(* IEC 61131-3 sources: daoli-st-library/DL_Process (part 65) *)

(* ---- FB_DL_EnthalpyCompareCtrl.st ---- *)
(*==============================================================================
 * 组件名称 (Component)  : FB_DL_EnthalpyCompareCtrl
 * 所属子库 (Sublibrary) : DL_Process
 * 当前版本 (Version)    : 1.0.1
 * 组件分类 (Category)   : 功能块（FUNCTION_BLOCK）· 焓差经济器比较控制 ·
 *                         Level 2 行业池 9.5 节 P0 链路闭环示范
 * 兼容性   (Platform)   : CODESYS 3.5 / TwinCAT 3 / 汇川 InoProShop / Schneider
 *                         Machine Expert；仅依赖 Standard.library 与本库已入库
 *                         算法函数，零厂商方言
 * 功能描述 (Function)   : 焓差比较控制执行块。新风/回风温湿度 4 输入 → 每拍
 *                         两次调用 FC_DL_HumidAirEnthalpy 计算双侧比焓 →
 *                         差分焓值判据（施密特迟滞防临界抖动）→ 新风阀位指令
 *                         输出；含最小新风位硬下限（卫生通风底线）与 ASHRAE
 *                         90.1 新风焓值高限停机语义（回差=死区防振荡）。
 *
 * 【干球温度判据陷阱警示 / Dry-bulb trap warning】
 *   本块判据【只允许使用焓差】，严禁以干球温差（fOaTempC 与 fRaTempC 比较）
 *   代替焓差判据：湿工况下新风干球温度可以低于回风，但其潜热（含湿量）更高，
 *   总焓反而高于回风——若按干球降温直觉开大新风阀，会引入高焓湿空气增加表冷
 *   负荷（验收向量 V1 复现此陷阱）。任何把本块改为干球比较的改动均视为破坏
 *   焓差经济器物理语义。
 *
 * 设计要点 (Key notes)  : ① 连续量组件 → 设 bInit 首扫（R19 唯一合法范式
 *                           IF bTrack OR (NOT bInit)），首扫输出最小新风位
 *                           安全值并重建迟滞态，运行中途 bTrack 一拍即重同步；
 *                         ② 迟滞状态机：开侧 fOaEnth < fRaEnth − 死区、关侧
 *                           fOaEnth > fRaEnth + 死区，死区区间内保持原态
 *                           （传感器漂移防线）；CASE + ELSE 非法态兜底；
 *                         ③ 高限停机：fEnthalpyHighLimit > 0 使能，fOaEnth
 *                           ≥ 高限 → 停机锁 bHighLimitTrip，回落至
 *                           高限 − 死区 以下才解除（瞬时型每拍重算，R15）；
 *                         ④ 失效语义（R11 裁定 D2）：任一温湿度/大气压非有
 *                           限值或越出引脚域 → 阀位指令输出最小新风位（安全
 *                           侧兜底），fOaEnthalpy/fRaEnthalpy/bHighLimitTrip
 *                           冻结保持末次有效值（诊断量冻结），故障码锁存，
 *                           仅「输入恢复 + bReset 上升沿」解除（R15）；
 *                         ⑤ 时间/温湿度全部引脚注入，禁读 CPU 本地钟；
 *                         ⑥ 限幅域对调自修复：fMinOaPos > fFreeCoolOaPos
 *                           时对调继续计算（公约 0.6），量纲注释与限幅域一致。
 * 枚举归属 (Enum note)  : E_DL_EnthalpyHyst（迟滞双侧态）随本块同文件发布；
 *                         本块不重复声明任何既有枚举。
 * 依赖     (Depends)    : FC_DL_HumidAirEnthalpy（DL_Algo，公开接口直接调用，
 *                         不内联重实现其焓值公式）；Standard.library
 *                         （R_TRIG / ABS / MIN / MAX / LIMIT）。
 * 开源溯源 (Origin)     : 原创实现（参考 ASHRAE 90.1 economizer 高限判据与
 *                         OSCAT Building 焓差经济器行为定义，clean-room）。
 *                         仅借鉴公开判据语义（差分焓值切换、最小新风位底线、
 *                         高限停机），未读取、未复制任何源码行；迟滞状态机、
 *                         失效冻结语义与码表为本库独立设计。
 * 故障码表 (Error codes):
 *   16#0005_0202【故障级】焓值计算输入失效（非有限值/越引脚域，锁存，
 *                 解除条件：输入恢复 AND bReset 上升沿）
 *   16#0005_0201【故障级】非法状态兜底（CASE ELSE，复用本库既有同义码，
 *                 与 FB_DL_PackMlStateMachine 同语义，公共码先例
 *                 DL_Algo 16#0002_0004）
 *   16#0005_0103【信息级】下游算法函数钳位码透传归并（温度/湿度/大气压
 *                 越界已钳位照算）/ 限幅域对调自修复（公约 0.6，本块唯一
 *                 分配信息级码复用，见 R11 D3）
 * 【规格偏离留档 / R11 Deviation register】
 *   D1 规格分配故障码 0005_0201（输入失效）与子库既有台账冲突（0201 已被
 *      R5 PackML 非法状态兜底占用）：按公约 0.7 冲突顺延，输入失效改用
 *      0005_0202；非法状态兜底与规格 0005_0202 分配冲突 → 复用既有同义码
 *      0005_0201。语义不变，仅码位重排。
 *   D2 规格失效语义同时出现「冻结保持末次有效阀位」与「输出 fMinOaPos 兜
 *      底值」：裁定为阀位指令输出 fMinOaPos（安全侧），焓值诊断输出与高限
 *      锁存位冻结末次有效值。
 *   D3 限幅域对调自修复（公约 0.6）码位：本块仅分配信息级 0005_0103，对调
 *      事件与下游钳位透传共用该码（当拍 uErrorId 择一呈现，均为信息级）。
 *   D4 新风干球负温域（-30..0 摄氏度）超出下游焓值函数计算域（0..100）：
 *      负干球工况下游返回 0 摄氏度钳位焓值（对新风焓偏高估计 → 判据偏保守
 *      安全侧），钳位信息经 0005_0103 当拍呈现；是否放行负干球工况由调用方
 *      按 D4 取舍（本块按引脚域 -30..60 验收输入，不自行拒绝）。
 * 红线自检 (Redline)    : R1 ✓ 零全局变量表与外部变量引用 ｜ R2 ✓ 零物理 IO 地址直写
 *                         R3 ✓ 纯 IEC 61131-3 ｜ R4 ✓ 非有限值防御（fX<>fX 先检再比较）
 *                             +迟滞判据浮点禁判等+本块无除法运算
 *                         R5 ✓ 全变量中英双语同行注释 ｜ R6 ✓ 迟滞状态机 ENUM+CASE
 *                             且 CASE-ELSE 兜底（码 0005_0201）
 *                         R7 ✓ R_TRIG 实例主体无条件周期刷新（严禁入分支）
 * 修订历史 (Revision)   :
 *   2026-11-15  v1.0.0  首版入库 · Round 06 · 泳道 C · 契约出处 ROUND_PLAN_R6 §3.14
 *   2026-11-15  v1.0.1  终审修复【工程语义级】参数 REAL 输入非数防御缺口：
 *                       原实现仅防御 5 个过程输入，fMinOaPos/fFreeCoolOaPos
 *                       非数经 LIMIT 直透生效域并输出 NaN 阀位指令（无故障
 *                       码伴随）；fEnthalpyDeadband 非数使迟滞判据恒 FALSE
 *                       冻结；fEnthalpyHighLimit 补显式自比检测。另阀位对
 *                       调改为经中间变量交换已防御生效值（防原始引脚穿透，
 *                       与 FB_DL_AnalogValve 终审修复同型）。修法遵循 R4
 *                       #15 沉淀范式：全部 REAL 输入（含参数）非数先检。
 *                       引脚契约零变更。
 * 验收向量 (Acceptance) :
 *   V1 干球陷阱：Oa=20.0 摄氏度/90.0%（焓≈53.6）vs Ra=26.0 摄氏度/40.0%
 *      （焓≈47.5）——新风干球低 6 摄氏度但焓高 6.1，判据不开经济器
 *      （bEconomizerActive=FALSE，阀位=最小新风位）；若按干球比较将错误开阀
 *   V2 迟滞往返：Oa=18.0/50.0（焓≈34.3）vs Ra=26.0/40.0（焓≈47.5），差
 *      −13.2 < −死区 2.0 → 开侧；Oa 渐升至 21.0/70.0（焓≈48.8），差 +1.0
 *      落在 ±2.0 死区内 → 保持开侧不抖动；Oa=22.0/75.0（焓≈53.7），差
 *      +5.9 > +2.0 → 关侧
 *   V3 高限停机：fEnthalpyHighLimit=60.0，Oa 焓 63.0 → bHighLimitTrip=TRUE
 *      强制最小新风位；Oa 焓回落至 58.0（< 60−2）才解除（回差防振荡）
 *   V4 硬下限：fMinOaPos=30.0 / fFreeCoolOaPos=100.0，任意路径断言
 *      fOaDamperCmd ≥ 30.0（激活 100.0 / 非激活 30.0）
 *   V5 非有限值冻结：fOaTempC 注入 NaN → 0005_0202 锁存、阀位回 fMinOaPos、
 *      焓值输出冻结末次有效值；输入恢复 + bReset 沿 → 清码恢复计算
 *   V6 中途 bTrack：运行中（开侧）注入 bTrack 一拍 → 迟滞重建为关侧、
 *      阀位回 fMinOaPos（R19 必测，不锁死）
 *============================================================================*)

(*-----------------------------------------------------------------------------
 * 调用示例 (Instance guide)：
 *   fbEco.fOaTempC := stMet.fTemp;          // 新风温湿度（滤波后信号）
 *   fbEco.fOaRelHum := stMet.fRh;
 *   fbEco.fRaTempC := stZone.fTemp;         // 回风/室内温湿度
 *   fbEco.fRaRelHum := stZone.fRh;
 *   fbEco.fEnthalpyHighLimit := 60.0;       // 0 = 禁用高限停机
 *   fbEco(bEnableCooling := bChwDemand,     // 周期调用
 *         bTrack := bHmiResync, bReset := bFaultReset);
 *   阀执行层（调用方职责）：fOaDamperCmd 直驱新风阀，下限保证亦由执行层
 *   复核；bHighLimitTrip 可联动压缩机保护。bTrack 用于 HMI 强制重同步。
 *----------------------------------------------------------------------------*)

{attribute 'qualified_only'}
{attribute 'strict'}
TYPE E_DL_EnthalpyHyst :
(
    eClosed := 0,   // 迟滞关侧：经济器停用，阀位=最小新风位（Closed side: economizer off, damper at minimum position）
    eOpened := 10   // 迟滞开侧：经济器激活，阀位=经济器全开位（Opened side: economizer active, damper at free-cooling position）
) UINT;
END_TYPE

FUNCTION_BLOCK FB_DL_EnthalpyCompareCtrl
VAR_INPUT
    fOaTempC           : REAL;             // 新风干球温度（Outdoor air dry-bulb temp）[摄氏度] 有效域 -30..60，越域按输入失效处理
    fOaRelHum          : REAL;             // 新风相对湿度（Outdoor air relative humidity）[百分数] 有效域 1..100，越域按输入失效处理
    fRaTempC           : REAL;             // 回风干球温度（Return air dry-bulb temp）[摄氏度] 有效域 0..100（与焓值 FC 计算域一致），越域按输入失效处理
    fRaRelHum          : REAL;             // 回风相对湿度（Return air relative humidity）[百分数] 有效域 1..100
    fAtmPress          : REAL := 101.325;  // 大气压（Atmospheric pressure）[kPa] 默认标准大气，透传焓值 FC，非有限值按输入失效处理
    fEnthalpyDeadband  : REAL := 2.0;      // 焓差切换死区（Enthalpy changeover deadband）[kJ/kg] 施密特迟滞半宽，默认 2.0，负值防御钳位为 0
    fMinOaPos          : REAL := 30.0;     // 最小新风阀位（Minimum outdoor air damper position）[百分数] 卫生通风硬下限，默认 30.0，域 0..100
    fFreeCoolOaPos     : REAL := 100.0;    // 经济器全开阀位（Free-cooling damper position）[百分数] 默认 100.0，域 0..100
    fEnthalpyHighLimit : REAL := 0.0;      // 新风焓值高限停机门限（Enthalpy high-limit trip）[kJ/kg] 默认 0=禁用（ASHRAE 90.1 高限语义）
    bEnableCooling     : BOOL := FALSE;    // 供冷需求使能（Cooling demand enable）[1] FALSE 时阀位恒回最小新风位
    bReset             : BOOL := FALSE;    // 复位（Reset）[1] 上升沿：输入失效锁存码仅在输入已恢复且本沿到达时清除
    bTrack             : BOOL := FALSE;    // 跟踪重同步（Track resync）[1] TRUE 时阀位回最小新风位并重建迟滞态（R19 必测）
END_VAR
VAR_OUTPUT
    fOaEnthalpy        : REAL;             // 新风比焓（Outdoor air enthalpy）[kJ/kg 干空气] 供 HMI/诊断；输入失效拍冻结末次有效值
    fRaEnthalpy        : REAL;             // 回风比焓（Return air enthalpy）[kJ/kg 干空气] 输入失效拍冻结末次有效值
    bEconomizerActive  : BOOL;             // 经济器激活（Economizer active）[1] 差分焓值判据通过且迟滞态为开侧
    fOaDamperCmd       : REAL;             // 新风阀位指令（Outdoor air damper command）[百分数] 量纲=阀位域 0..100，硬下限恒 ≥ fMinOaPos
    bHighLimitTrip     : BOOL;             // 焓值高限停机（Enthalpy high-limit trip）[1] 激活中；失效拍冻结末次有效值
    uErrorId           : UDINT;            // 事件码（Error code）16#0005_0202 输入失效（锁存）/ 16#0005_0201 非法态兜底 / 16#0005_0103 信息级；0 = 无
END_VAR
VAR
    bInit              : BOOL := FALSE;    // 首扫标志（First-scan flag，R19 范式配套）
    _eHyst             : E_DL_EnthalpyHyst := E_DL_EnthalpyHyst.eClosed;  // 迟滞状态机内部态（Internal hysteresis state）
    _bFailLatch        : BOOL := FALSE;    // 输入失效锁存（Input-failure latch，仅解除路径清码 R15）
    _bInFailNow        : BOOL;             // 本拍输入失效判定（Input failure this scan，瞬时条件）
    _bOaTOk            : BOOL;             // 新风温度有效（OA temp valid）
    _bOaROk            : BOOL;             // 新风湿度有效（OA humidity valid）
    _bRaTOk            : BOOL;             // 回风温度有效（RA temp valid）
    _bRaROk            : BOOL;             // 回风湿度有效（RA humidity valid）
    _bPOk              : BOOL;             // 大气压有限（Pressure finite）
    _bClampInfo        : BOOL;             // 下游钳位信息标志（Downstream clamp info flag，当拍）
    _bSwapInfo         : BOOL;             // 限幅域对调标志（Span-swap repair flag，公约 0.6，当拍）
    _bElseHit          : BOOL;             // 非法态兜底命中标志（Illegal-state fallback hit，当拍）
    fDbC               : REAL;             // 生效死区（Effective deadband）[kJ/kg] 负值钳位为 0 后
    fMinPosC           : REAL;             // 生效最小新风位（Effective min position）[百分数] 钳位域 0..100
    fCoolPosC          : REAL;             // 生效全开阀位（Effective free-cool position）[百分数] 钳位域 0..100
    fPosTmp            : REAL;             // 阀位对调交换中间变量（Damper swap temp carrier）[百分数]，生效域已防御值
    uErrOa             : UDINT;            // 新风焓值 FC 返回码（OA enthalpy FC code）
    uErrRa             : UDINT;            // 回风焓值 FC 返回码（RA enthalpy FC code）
    fbTrigReset        : R_TRIG;           // 复位信号上升沿检测实例（Reset edge detector）
END_VAR
VAR CONSTANT
    DL_ENT_INF_MAX     : REAL := 1.0E30;   // 有限值判定幅值上限（Magnitude bound for finite-value check）
    DL_ENT_OA_T_MIN    : REAL := -30.0;    // 新风温度验收域下限（OA temp domain floor）[摄氏度]
    DL_ENT_OA_T_MAX    : REAL := 60.0;     // 新风温度验收域上限（OA temp domain ceiling）[摄氏度]
    DL_ENT_RA_T_MIN    : REAL := 0.0;      // 回风温度验收域下限=焓值 FC 计算域下限（RA temp domain floor）[摄氏度]
    DL_ENT_RA_T_MAX    : REAL := 100.0;    // 回风温度验收域上限=焓值 FC 计算域上限（RA temp domain ceiling）[摄氏度]
    DL_ENT_RH_MIN      : REAL := 1.0;      // 湿度验收域下限（Humidity domain floor）[百分数]
    DL_ENT_RH_MAX      : REAL := 100.0;    // 湿度验收域上限（Humidity domain ceiling）[百分数]
    DL_ENT_POS_MIN     : REAL := 0.0;      // 阀位域下限（Damper domain floor）[百分数]
    DL_ENT_POS_MAX     : REAL := 100.0;    // 阀位域上限（Damper domain ceiling）[百分数]
END_VAR

// -----------------------------------------------------------------------------
// 段 1｜复位沿实例无条件周期刷新（R7 红线：严禁移入 IF/CASE 分支）
// -----------------------------------------------------------------------------
fbTrigReset(CLK := bReset);                 // 复位沿检测

// -----------------------------------------------------------------------------
// 段 2｜出口默认值与参数防御准备（公约 0.8：默认值先于防御路径；0.6 对调自修复）
// -----------------------------------------------------------------------------
uErrorId := 16#0000_0000;                   // 事件码先清零（后续按优先级覆盖）
_bClampInfo := FALSE;                       // 钳位信息标志每拍重算
_bSwapInfo := FALSE;                        // 对调标志每拍重算
_bElseHit := FALSE;                         // 兜底命中标志每拍重算
bEconomizerActive := FALSE;                 // 经济器指示默认停用（迟滞段重判）

fDbC := fEnthalpyDeadband;                  // 死区原值生效
IF fDbC <> fDbC THEN
    fDbC := 2.0;                            // 非数防御（公约 0.8 参数全覆盖，终审修复）：回落默认死区
END_IF
IF fDbC < 0.0 THEN
    fDbC := 0.0;                            // 防御钳位：负死区无物理意义，按 0（无迟滞）处理
END_IF

fMinPosC := fMinOaPos;                      // 最小新风位先做非数防御再钳位（终审修复）
IF fMinPosC <> fMinPosC THEN
    fMinPosC := 30.0;                       // 非数回落默认最小新风位 [百分数]
END_IF
fMinPosC := LIMIT(DL_ENT_POS_MIN, fMinPosC, DL_ENT_POS_MAX);      // 最小新风位钳位 [百分数]
fCoolPosC := fFreeCoolOaPos;                // 全开阀位先做非数防御再钳位（终审修复）
IF fCoolPosC <> fCoolPosC THEN
    fCoolPosC := 100.0;                     // 非数回落默认全开阀位 [百分数]
END_IF
fCoolPosC := LIMIT(DL_ENT_POS_MIN, fCoolPosC, DL_ENT_POS_MAX);    // 全开阀位钳位 [百分数]
IF fMinPosC > fCoolPosC THEN
    fPosTmp   := fMinPosC;                  // 对调经已防御生效值交换（中间变量，防原始引脚
    fMinPosC  := fCoolPosC;                 // 非有限值穿透回生效域，终审修复）
    fCoolPosC := fPosTmp;                   // 对调后半程
    _bSwapInfo := TRUE;                     // 对调事件置信息级标志（码 0005_0103，R11 D3）
END_IF

// -----------------------------------------------------------------------------
// 段 3｜R19 首扫/跟踪同步：判据唯一合法范式 IF bTrack OR (NOT bInit)
//       首扫输出最小新风位安全值；运行中途跟踪脉冲重建迟滞态不锁死（验收 V6）
// -----------------------------------------------------------------------------
IF bTrack OR (NOT bInit) THEN
    _eHyst := E_DL_EnthalpyHyst.eClosed;    // 迟滞态重建为关侧
    bEconomizerActive := FALSE;             // 经济器指示停用
    bHighLimitTrip := FALSE;                // 高限锁存重建
    fOaDamperCmd := fMinPosC;               // 首扫/跟踪安全值：最小新风位 [百分数]
    bInit := TRUE;                          // 首扫完成
END_IF

// -----------------------------------------------------------------------------
// 段 4｜输入有效性防御（公约 0.8：全部 REAL 输入先做 fX<>fX 检测再比较）
// -----------------------------------------------------------------------------
_bOaTOk := (NOT (fOaTempC <> fOaTempC)) AND (ABS(fOaTempC) <= DL_ENT_INF_MAX)
       AND (fOaTempC >= DL_ENT_OA_T_MIN) AND (fOaTempC <= DL_ENT_OA_T_MAX);      // 新风温度：非有限值 + 引脚域
_bOaROk := (NOT (fOaRelHum <> fOaRelHum)) AND (ABS(fOaRelHum) <= DL_ENT_INF_MAX)
       AND (fOaRelHum >= DL_ENT_RH_MIN) AND (fOaRelHum <= DL_ENT_RH_MAX);        // 新风湿度：非有限值 + 域
_bRaTOk := (NOT (fRaTempC <> fRaTempC)) AND (ABS(fRaTempC) <= DL_ENT_INF_MAX)
       AND (fRaTempC >= DL_ENT_RA_T_MIN) AND (fRaTempC <= DL_ENT_RA_T_MAX);      // 回风温度：非有限值 + 域
_bRaROk := (NOT (fRaRelHum <> fRaRelHum)) AND (ABS(fRaRelHum) <= DL_ENT_INF_MAX)
       AND (fRaRelHum >= DL_ENT_RH_MIN) AND (fRaRelHum <= DL_ENT_RH_MAX);        // 回风湿度：非有限值 + 域
_bPOk := (NOT (fAtmPress <> fAtmPress)) AND (ABS(fAtmPress) <= DL_ENT_INF_MAX);   // 大气压：仅非有限值防御（域由下游钳位）
_bInFailNow := NOT (_bOaTOk AND _bOaROk AND _bRaTOk AND _bRaROk AND _bPOk);       // 任一失效即本拍失效

// -----------------------------------------------------------------------------
// 段 5｜失效锁存（R15：锁存型只在解除路径清码——输入恢复 AND 复位沿）
// -----------------------------------------------------------------------------
IF _bInFailNow THEN
    _bFailLatch := TRUE;                    // 失效条件置位锁存
END_IF
IF fbTrigReset.Q AND (NOT _bInFailNow) THEN
    _bFailLatch := FALSE;                   // 解除路径：输入已恢复 + 复位沿
END_IF

// -----------------------------------------------------------------------------
// 段 6｜失效路径：安全侧兜底输出 + 诊断量冻结（R11 D2 裁定语义）
//       阀位指令回最小新风位；焓值/高限位保持末次有效值（FB 输出静态保持，
//       非未初始化路径，出口确定）
// -----------------------------------------------------------------------------
IF _bFailLatch THEN
    uErrorId := 16#0005_0202;               // 输入失效【故障级】（顺延码位，R11 D1）
    bEconomizerActive := FALSE;             // 安全侧：经济器停用
    _eHyst := E_DL_EnthalpyHyst.eClosed;    // 恢复后迟滞从关侧重建
    fOaDamperCmd := fMinPosC;               // 阀位兜底：最小新风位 [百分数]
    // fOaEnthalpy / fRaEnthalpy / bHighLimitTrip 不赋值 = 冻结末次有效值
ELSE

    // -------------------------------------------------------------------------
    // 段 7｜焓值计算：每拍两次调用 FC_DL_HumidAirEnthalpy（公开接口直接调用，
    //       禁止内联重实现其公式链）
    // -------------------------------------------------------------------------
    uErrOa := 16#0000_0000;                 // 返回码先清零
    uErrRa := 16#0000_0000;                 // 返回码先清零
    fOaEnthalpy := FC_DL_HumidAirEnthalpy(fTempC := fOaTempC, fRelHum := fOaRelHum,
                                          fAtmPress := fAtmPress, uErrorId => uErrOa);  // 新风比焓 [kJ/kg 干空气]
    fRaEnthalpy := FC_DL_HumidAirEnthalpy(fTempC := fRaTempC, fRelHum := fRaRelHum,
                                          fAtmPress := fAtmPress, uErrorId => uErrRa);  // 回风比焓 [kJ/kg 干空气]

    // 双调用返回码并集归并（0.8 防御兜底：下游拒绝码理论上段 4 已拦截）
    IF (uErrOa = 16#0002_0004) OR (uErrRa = 16#0002_0004) THEN
        _bFailLatch := TRUE;                // 下游拒绝 → 转入失效锁存（下一拍走段 6）
        uErrorId := 16#0005_0202;           // 输入失效【故障级】
        bEconomizerActive := FALSE;         // 安全侧停用
        fOaDamperCmd := fMinPosC;           // 阀位兜底 [百分数]
    ELSE
        _bClampInfo := (uErrOa <> 16#0000_0000) OR (uErrRa <> 16#0000_0000);
                                            // 任一钳位码（1701/1702/1703）→ 信息级透传归并（R11 D4）

        // ---------------------------------------------------------------------
        // 段 8｜高限停机（ASHRAE 90.1 语义）：瞬时型每拍重算 + 死区回差防振荡
        //       （R15：非锁存位，激活条件存在即呈现，回差内保持）
        // ---------------------------------------------------------------------
        IF (fEnthalpyHighLimit = fEnthalpyHighLimit) AND (fEnthalpyHighLimit > 0.0) THEN
            // 非数门限按禁用处理（公约 0.8 显式检测，终审修复：NaN 比较恒 FALSE
            // 虽天然落入禁用分支，仍显式自比检测防方言差异）
            IF fOaEnthalpy >= fEnthalpyHighLimit THEN
                bHighLimitTrip := TRUE;     // 新风焓达高限 → 停机锁激活
            ELSIF fOaEnthalpy < (fEnthalpyHighLimit - fDbC) THEN
                bHighLimitTrip := FALSE;    // 回落至回差下界之下才解除
            END_IF                          // 回差区间内保持原态（防临界振荡）
        ELSE
            bHighLimitTrip := FALSE;        // 门限 0 = 高限停机禁用
        END_IF

        // ---------------------------------------------------------------------
        // 段 9｜差分焓值迟滞状态机（ENUM + CASE + ELSE 兜底，红线 R6）
        //       【干球陷阱警示】此处只允许焓差比较，严禁改为干球温差判据
        // ---------------------------------------------------------------------
        CASE _eHyst OF

            E_DL_EnthalpyHyst.eClosed:      // 关侧：等待开侧判据
                IF bEnableCooling AND (NOT bHighLimitTrip)
                   AND (fOaEnthalpy < fRaEnthalpy - fDbC) THEN
                    _eHyst := E_DL_EnthalpyHyst.eOpened;   // 新风焓显著低于回风 → 开侧
                END_IF

            E_DL_EnthalpyHyst.eOpened:      // 开侧：等待关侧判据或退出条件
                IF (NOT bEnableCooling) OR bHighLimitTrip
                   OR (fOaEnthalpy > fRaEnthalpy + fDbC) THEN
                    _eHyst := E_DL_EnthalpyHyst.eClosed;   // 退出条件任一 → 关侧
                END_IF

            ELSE                            // 非法状态兜底（故障级 0005_0201）
                _bElseHit := TRUE;          // 当拍呈现码
                _eHyst := E_DL_EnthalpyHyst.eClosed;       // 回关侧安全态
        END_CASE

        // ---------------------------------------------------------------------
        // 段 10｜输出合成：经济器指示 + 阀位指令（最小新风硬下限双保险）
        // ---------------------------------------------------------------------
        bEconomizerActive := (_eHyst = E_DL_EnthalpyHyst.eOpened);  // 判据通过且迟滞态为开侧
        IF bEconomizerActive THEN
            fOaDamperCmd := fCoolPosC;      // 激活：经济器全开位 [百分数]
        ELSE
            fOaDamperCmd := fMinPosC;       // 非激活：最小新风位 [百分数]
        END_IF
        fOaDamperCmd := MAX(fOaDamperCmd, fMinPosC);   // 硬下限出口断言（对调后恒真，双保险）

        // ---------------------------------------------------------------------
        // 段 11｜事件码优先级合成（R21：信息级只进 uErrorId）：兜底 > 信息级 > 无
        // ---------------------------------------------------------------------
        IF _bElseHit THEN
            uErrorId := 16#0005_0201;       // 非法状态兜底【故障级】（复用同义码，R11 D1）
        ELSIF _bClampInfo OR _bSwapInfo THEN
            uErrorId := 16#0005_0103;       // 下游钳位透传 / 限幅域对调【信息级】
        END_IF                              // 否则保持段 2 清零值
    END_IF
END_IF

END_FUNCTION_BLOCK

(* ---- FB_DL_EscHeLeakCheck.st ---- *)
(*==============================================================================
 * 组件名称 (Component)  : FB_DL_EscHeLeakCheck
 * 所属子库 (Sublibrary) : DL_Process
 * 当前版本 (Version)    : 1.0.1
 * 组件分类 (Category)   : 功能块（FUNCTION_BLOCK）· 静电吸盘氦背冷泄漏率判定
 * 兼容性   (Platform)   : CODESYS 3.5 / TwinCAT 3 / 汇川 InoProShop / Schneider Machine Expert
 *                         仅依赖 Standard.library（R_TRIG / TON / ABS / MIN / MAX / LIMIT），零厂商方言
 * 接口依赖 (Depends)    : E_DL_Ne107Status —— 唯一属主为 DL_Device 子库的契约件
 *                         I_DL_DeviceHealth（R13 泳道 A1）。本文件只引用成员，不重定义枚举体。
 * 功能描述 (Function)   : 静电吸盘（ESC）氦背冷回路的三段式泄漏率判定 ——
 *                         升压段（斜率监视 + 达压确认）→ 稳压段（窗内极差稳定判据）→
 *                         测量段（压降率 → 漏率换算 + 温漂修正）→ 判定（OK / Warn / NG）。
 * 与 FB_DL_LeakTestStation 的分工（必须遵守，禁止合并）:
 *                         后者是**通用压降法工站**（充气-稳压-保压-压降换算-排气，面向工件
 *                         腔体，压力区间宽、带排气相与夹具确认）；本件是**ESC 专用**：氦侧
 *                         压力区间窄（1~100 kPa）、必须做温漂修正、判定带 Warn 三级、且要
 *                         单独识别「氦源串漏方向」（测量段压力上升 = 阀未关或源侧串漏）。
 *                         两者**不得合并**：合并会把两套压力量纲与判定门限塞进一个方式参数，
 *                         这正是历史库反复交学费的老毛病（一套 MODE 管两种物理过程）。
 * 边界     (Boundary)   : ① 不做抽真空/排气相（ESC 背冷不排气，氦侧常压回收）；② 不做
 *                         夹具确认（背冷腔由卡盘机械结构保证）；③ 不做腔体几何漏率模型，
 *                         压降率→漏率的换算系数为标定常量（见 DL_ESC_LEAK_K 注释）。
 * 分层声明 (Layer)      : 工艺层（DL_Process）。零全局变量表引用、零外部变量声明、零物理 IO。
 * 段序     (Segments)   : 段1 实例无条件刷新 → 段2 断输入拍自清与复位通道（CASE 前，R39）→
 *                         段3 输入防御与参数钳位 → 段4 启动沿受理（R24/R25）→ 段5 相位状态机 →
 *                         段6 判定结算 → 段7 码位单一优先级链 → 段8 出口钳位与保持重写。
 * 枚举映射表 (R31)      : 相位 E_DL_EscLeakPhase：eIdle(0)→标签 0｜ePressurize(10)→标签 10｜
 *                         eStabilize(20)→标签 20｜eMeasure(30)→标签 30｜eVerdict(40)→标签 40｜
 *                         eFault(99)→标签 99。结果 E_DL_LeakResult：eOk(0)｜eWarn(10)｜
 *                         eNg(20)｜eAborted(30)，不作为 CASE 选择子，仅作出口判定值。
 * 单拍标志清单 (R25)    : bStart —— 预清零点：段1 每拍被实例输出覆盖；置位点：段1
 *                         `_bStartReq := _fbTrigStart.Q AND (NOT _bStartConsumed)`；自清点：
 *                         段4 消费时置 `_bStartConsumed := TRUE`，bStart 回 FALSE 即解除。
 *                         bReset —— 预清零点：段1 覆盖 _bResetEdge；置位点：段1 实例调用；
 *                         自清点：紧随实例调用的 _bResetEdge 赋值行。
 * 保持位清单 (R27)      : bDone / bPass / eResult / fLeakRate / fPressDecay —— 逐拍由
 *                         _bDoneLatched / _bPassLatched / _eResultHeld / _fLeakHeld /
 *                         _fDecayHeld 重写并夹域；新启动沿与复位沿清除。
 * 定时器清单 (R40)      : 三段各一个 TON，**每段切换必须断输入一拍**（R40 核心）：
 *                         _fbTonPress ｜IN = (相位 = ePressurize) AND NOT _bPressBreak｜
 *                         断输入标志 _bPressBreak（进升压段置一拍，段2 自清）；
 *                         _fbTonStab   ｜IN = (相位 = eStabilize) AND NOT _bStabBreak｜
 *                         断输入标志 _bStabBreak（进稳压段置一拍，段2 自清）；
 *                         _fbTonStabExt｜IN = (相位 = eStabilize) AND _bStabExtended AND NOT _bStabExtBreak｜
 *                         断输入标志 _bStabExtBreak（延长一次时置一拍，段2 自清）；
 *                         _fbTonMeas   ｜IN = (相位 = eMeasure) AND NOT _bMeasBreak｜
 *                         断输入标志 _bMeasBreak（进测量段置一拍，段2 自清）。
 *                         四者绝不共用实例、绝不用 `IN := (相位 <> eIdle)` 这类跨段恒真写法。
 * 三元一致表 (R35)      : 达压容差守卫 0.01~50 kPa / 封顶 50 / 判据 `≤`｜
 *                         漏率 Warn 阈守卫 0~1E4 sccm / 封顶 1E4 / 判据 `>`（超 Warn 进 Warn 带）｜
 *                         漏率 NG 阈守卫 0~1E4 sccm 且强制 ≥ Warn / 判据 `>`（超 NG 判 NG）。
 * 镜像量清单 (R38)      : fHePressure 的唯一消费点是段3 的 _fPnow（每拍单次锁存），相位机
 *                         与结算全部读 _fPnow，绝不回读实时入参；fChuckTemp 同理锁存为 _fTnow。
 * 开源溯源 (Origin)     : 自研（T2-8 仅借「分级 → 维护建议」的语言形态，即 Warn/NG 两级
 *                         判定后给出维护动作，不涉及任何实现细节）。ESC 氦背冷检漏无可对应
 *                         的开源件（LBP 与 OSCAT 均无此工艺块，见 R13 溯源结论），压降率→
 *                         漏率换算与三段定时结构为本库独立设计。许可证说明：无代码借鉴对象，
 *                         本文件为本库原创，随本库许可证发布。
 * 验收向量 (Acceptance) :
 *   V1 15 kPa 达压、30 s 内压降 0.04 kPa → fPressDecay ≈ 0.00133 kPa/s、
 *      fLeakRate ≈ 2.0 sccm（× 换算系数 1500）→ eOk、bPass = TRUE（保持）。
 *   V2 压降 0.12 kPa/30 s → 漏率 6.0 sccm > NG 阈 5.0 → eNg、bPass = FALSE（保持）。
 *   V3（V-C 三段定时器，R40）升压 10 s + 稳压 10 s + 测量 30 s，三段各用一个 TON 且
 *      **每段切换断输入一拍**。若误写成三段共用一个 TON 且 IN 跨段恒真，则 50 s 时
 *      tMeasure = 30 s 会被提前判超时 —— 本向量用于区分这两种实现。
 *   V4（V-D 中止恢复，R41）eMeasure 中 bEnable 掉 → 回 eIdle、eResult = eAborted、
 *      bDone 保持；重新 bStart 后三段计时**从 0 开始**（断输入拍保证 ET 清零）。
 *   V5（V-A 非有限）fHePressure = NaN → 16#0005_02F8、fLeakRate 保持上次值（绝不写 NaN）。
 * 偏离留档 (Deviation)  :
 *   ① 输入非有限值与「非法状态兜底」共用 16#0005_02F8：规格故障表只给 3 个故障码，
 *      而其验收向量 V5 明确要求 NaN 走 02F8，故按向量口径执行，不新增码位。
 *   ② fPressRiseMax 的语义裁定：规格命名为「升压速率上限」。氦侧有机械减压阀，超压风险
 *      不成立，因此本件不把它当拦截阈值，而是当作**升压段的供气健康基准**：升压速率
 *      持续（≥1 s）低于其 2 % 且远未达压时判供气异常 02F6。「上限语义不拦截」这一裁定
 *      在头注释声明，避免后人误以为漏实现了超速拦截。
 *   ③ 漏率换算系数 DL_ESC_LEAK_K = 1500 sccm/(kPa/s) 为标定常量：由背冷腔容积与标定
 *      工装决定，规格未给容积引脚；调用方按腔体台账整定（值误差只影响绝对量程，
 *      不影响 OK/Warn/NG 的判定结构）。
 *   ④ 稳压延长仅一次（01C8 语义）；延长后仍不稳则**进入测量**但在判定时把 eOk 降为
 *      eWarn（不确定性上升），绝不因稳定判据未过而丢弃整次检测。
 * 修订历史 (Revision)   :
 *   2026-11-15  v1.0.0  首版入库（Round 13 · 泳道 C · DL_Process 第 24 件）
 *   2026-11-16  v1.0.1  终审修复：稳压延长窗原实现「_fbTonStab.Q OR _fbTonStabExt.Q」
 *                       联合裁决，延长置位后主稳压定时器 IN 未断、Q 保持 TRUE，下一拍
 *                       即被提前判「延长后仍不稳」进测量，_fbTonStabExt 从未计时；改为以
 *                       _bStabExtended 区分两窗，延长窗仅由 _fbTonStabExt.Q 裁决（D-C4-1）
 *============================================================================*)

(*-----------------------------------------------------------------------------
 * 枚举: E_DL_EscLeakPhase（归属 FB_DL_EscHeLeakCheck，同文件发布）
 *----------------------------------------------------------------------------*)
TYPE E_DL_EscLeakPhase :
(
    eIdle       := 0,   // 空闲：等启动沿 / Idle, awaiting the start edge
    ePressurize := 10,  // 升压：等达压或超时 / Pressurise, awaiting the target or a timeout
    eStabilize  := 20,  // 稳压：等窗内极差收敛 / Stabilise, awaiting a settled pressure range
    eMeasure    := 30,  // 测量：隔离测压降 / Measure, isolated pressure-decay window
    eVerdict    := 40,  // 判定：结算一次后回空闲 / Verdict, settles once then returns to idle
    eFault      := 99   // 故障：锁存等复位 / Fault latched until reset
) UINT;
END_TYPE

(*-----------------------------------------------------------------------------
 * 枚举: E_DL_LeakResult（归属 FB_DL_EscHeLeakCheck，同文件发布）
 *----------------------------------------------------------------------------*)
TYPE E_DL_LeakResult :
(
    eOk      := 0,      // 合格：漏率低于 Warn 阈 / OK, leak rate below the warn limit
    eWarn    := 10,     // 警告：落在 Warn 带或稳定判据欠佳 / Warn, inside the warn band or weakly settled
    eNg      := 20,     // 不合格：漏率超 NG 阈 / Reject, leak rate above the reject limit
    eAborted := 30      // 中止：无结论（掉使能或复位）/ Aborted, no conclusion
) UINT;
END_TYPE

FUNCTION_BLOCK FB_DL_EscHeLeakCheck
VAR_INPUT
    bEnable        : BOOL;                  // 使能（Enable），FALSE = 中止当前检测并回空闲；复位通道不受其屏蔽 / Enable, FALSE aborts the check
    bReset         : BOOL;                  // 复位（Reset），上升沿清故障、结果与保持量 / Rising edge clears fault, result and held values
    bStart         : BOOL;                  // 启动一次检测（One-shot start），上升沿受理（R24）/ One-shot start, rising edge only
    fHePressure    : REAL;                  // 氦侧压力（Helium pressure）[kPa]，域 0~500 / Helium pressure [kPa], 0 to 500
    fHeFlow        : REAL;                  // 氦侧流量（Helium flow）[sccm]，域 0~5000，用于与漏率交叉校验 / Helium flow [sccm], used for the cross check
    fChuckTemp     : REAL;                  // 卡盘温度（Chuck temperature）[℃]，域 0~200，温漂修正用 / Chuck temperature [degC], used for the drift correction
    tPressurizeMax : TIME := T#20S;         // 升压段超时（Pressurise timeout），默认 20 s / Pressurise timeout, default 20 s
    tStabilize     : TIME := T#10S;         // 稳压段时长（Stabilisation time），默认 10 s / Stabilisation time, default 10 s
    tMeasure       : TIME := T#30S;         // 测量段时长（Measurement time），默认 30 s / Measurement time, default 30 s
    fPressTarget   : REAL := 15.0;          // 目标背压（Target back pressure）[kPa]，域 1~100 / Target back pressure [kPa]
    fPressTol      : REAL := 0.5;           // 达压容差（Pressure tolerance）[kPa]，域 0.01~50 / Pressure tolerance [kPa]
    fLeakWarn      : REAL := 3.0;           // 漏率 Warn 阈（Leak-rate warn limit）[sccm]，域 0~1E4 / Leak-rate warn limit [sccm]
    fLeakNg        : REAL := 5.0;           // 漏率 NG 阈（Leak-rate reject limit）[sccm]，域 0~1E4 且 ≥ Warn / Leak-rate reject limit [sccm]
    fPressRiseMax  : REAL := 2.0;           // 升压速率基准（Pressurise rate reference）[kPa/s]，域 0.01~100，偏离留档② / Pressurise rate reference [kPa/s]
    fTempCoeff     : REAL := 0.003;         // 压力温漂修正系数（Pressure temperature coefficient）[1/K]，域 −0.05~0.05 / Pressure temperature coefficient [1/K]
    fStabTol       : REAL := 0.2;           // 稳压判据：窗内极差上限（Stabilisation tolerance）[kPa]，域 0.001~50 / Stabilisation tolerance [kPa]
END_VAR

VAR_OUTPUT
    fLeakRate      : REAL;                  // 换算漏率（Corrected leak rate）[sccm]，温漂修正后，夹进 ≥0 / Corrected leak rate [sccm], clamped non-negative
    fPressDecay    : REAL;                  // 测量段压降率（Pressure decay rate）[kPa/s]，有符号，夹域 / Pressure decay rate [kPa/s], signed and clamped
    eResult        : E_DL_LeakResult;       // 判定结果（Result），保持语义（R27）/ Result, held until the next start
    bDone          : BOOL;                  // 检测完成（Done），保持语义（R27）/ Done, held
    bPass          : BOOL;                  // 合格（Pass），保持语义（R27）/ Pass, held
    nTestCount     : UDINT;                 // 检测次数（Test counter）[次] / Test counter [count]
    nNgCount       : UDINT;                 // 不合格次数（Reject counter）[次] / Reject counter [count]
    eHealth        : E_DL_Ne107Status;      // 健康态（NE107 health），引用属主 A1 的枚举 / NE107 health, owned by A1
    uDiagCode      : UDINT;                 // 诊断码（Diagnostic code），本拍单一优先级链输出 / Diagnostic code, single priority chain
    uErrorId       : UDINT;                 // 故障码（Error code），仅故障级码，0 = 无故障 / Fault-level code, 0 = no fault
    bError         : BOOL;                  // 故障标志（Error），仅故障级码置位（NG 属工件不良，不置位）/ TRUE only for fault-level codes
END_VAR

VAR
    _ePhase        : E_DL_EscLeakPhase := E_DL_EscLeakPhase.eIdle;  // 内部相位（Internal phase）/ Internal phase value
    _bStartReq     : BOOL;                  // 启动单拍请求（Start one-shot request）/ Start one-shot request
    _bStartConsumed : BOOL;                 // 启动已消费（Start consumed flag）/ Start consumed flag
    _bResetEdge    : BOOL;                  // 复位沿单拍标志（Reset one-shot flag）/ Reset one-shot flag
    _bPressBreak   : BOOL;                  // 升压段断输入拍（Pressurise break）/ Pressurise segment break
    _bStabBreak    : BOOL;                  // 稳压段断输入拍（Stabilise break）/ Stabilise segment break
    _bStabExtBreak : BOOL;                  // 稳压延长段断输入拍（Stabilise extension break）/ Stabilise extension break
    _bMeasBreak    : BOOL;                  // 测量段断输入拍（Measure break）/ Measure segment break
    _uFaultCode    : UDINT;                 // 本拍故障级码（Fault-level code this scan）/ Fault-level code of this scan
    _uFaultLatched : UDINT;                 // 故障码锁存（Latched fault code），仅复位清除 / Latched fault code, reset only
    _uInfoCode     : UDINT;                 // 本拍信息级码（Info-level code this scan）/ Info-level code of this scan
    _bFaultCond    : BOOL;                  // 故障条件（Fault condition）/ Fault condition flag
    _fPnow         : REAL;                  // 压力快照（Pressure snapshot）[kPa]，唯一消费点的入口（R38）/ Pressure snapshot [kPa]
    _fTnow         : REAL;                  // 温度快照（Temperature snapshot）[℃]，唯一消费点的入口（R38）/ Temperature snapshot [degC]
    _fFlowNow      : REAL;                  // 流量快照（Flow snapshot）[sccm]，交叉校验用 / Flow snapshot [sccm]
    _fTargetEff    : REAL;                  // 生效目标压力（Effective target pressure）[kPa] / Effective target pressure [kPa]
    _fTolEff       : REAL;                  // 生效达压容差（Effective tolerance）[kPa] / Effective pressure tolerance [kPa]
    _fWarnEff      : REAL;                  // 生效 Warn 阈（Effective warn limit）[sccm] / Effective warn limit [sccm]
    _fNgEff        : REAL;                  // 生效 NG 阈（Effective reject limit）[sccm] / Effective reject limit [sccm]
    _fRiseRefEff   : REAL;                  // 生效升压速率基准（Effective rate reference）[kPa/s] / Effective rate reference [kPa/s]
    _fCoeffEff     : REAL;                  // 生效温漂系数（Effective temperature coefficient）[1/K] / Effective coefficient [1/K]
    _fStabTolEff   : REAL;                  // 生效稳压容差（Effective stabilisation tolerance）[kPa] / Effective tolerance [kPa]
    _fP0           : REAL;                  // 升压起点压力（Pressure at pressurise start）[kPa] / Pressure at pressurise start [kPa]
    _fPm           : REAL;                  // 测量起点压力（Pressure at measure start）[kPa] / Pressure at measure start [kPa]
    _fTm           : REAL;                  // 测量起点温度（Temperature at measure start）[℃] / Temperature at measure start [degC]
    _fStabMin      : REAL;                  // 稳压段压力极小（Stabilise minimum pressure）[kPa] / Stabilise minimum [kPa]
    _fStabMax      : REAL;                  // 稳压段压力极大（Stabilise maximum pressure）[kPa] / Stabilise maximum [kPa]
    _fStabRange    : REAL;                  // 稳压段极差（Stabilise range）[kPa] / Stabilise range [kPa]
    _bStabExtended : BOOL;                  // 稳压已延长（Stabilisation extended once）/ Stabilisation extended once
    _bStabWeak     : BOOL;                  // 稳定判据欠佳（Weakly settled）/ Weakly settled flag
    _fRiseRate     : REAL;                  // 升压速率（Pressurise rate）[kPa/s] / Pressurise rate [kPa/s]
    _fEtSec        : REAL;                  // 定时器已历秒值（Elapsed seconds）[s] / Elapsed seconds
    _fDecay        : REAL;                  // 压降量（Pressure drop）[kPa]，有符号 / Pressure drop [kPa], signed
    _fDecayCorr    : REAL;                  // 温漂修正后压降（Drift-corrected drop）[kPa] / Drift-corrected pressure drop [kPa]
    _fDecayRate    : REAL;                  // 压降率（Decay rate）[kPa/s] / Decay rate [kPa/s]
    _fMeasSec      : REAL;                  // 测量段实际秒值（Measured seconds）[s] / Measured seconds [s]
    _fLeakCalc     : REAL;                  // 本拍漏率（Computed leak rate）[sccm] / Computed leak rate [sccm]
    _fDtKelvin     : REAL;                  // 测量段温差（Temperature change）[K] / Temperature change during measure [K]
    _eResultCalc   : E_DL_LeakResult;       // 本拍结果（Computed result）/ Computed result
    _bDoneLatched  : BOOL;                  // 完成锁存（Done latch）/ Done latch
    _bPassLatched  : BOOL;                  // 合格锁存（Pass latch）/ Pass latch
    _eResultHeld   : E_DL_LeakResult := E_DL_LeakResult.eAborted;   // 保持的结果（Held result）/ Held result
    _fLeakHeld     : REAL;                  // 保持的漏率（Held leak rate）[sccm] / Held leak rate [sccm]
    _fDecayHeld    : REAL;                  // 保持的压降率（Held decay rate）[kPa/s] / Held decay rate [kPa/s]
    _nTestInt      : UDINT;                 // 内部检测计数（Internal test counter）[次] / Internal test counter [count]
    _nNgInt        : UDINT;                 // 内部不合格计数（Internal reject counter）[次] / Internal reject counter [count]
    _fbTrigStart   : R_TRIG;                // 启动上升沿（Start rising edge）/ Start rising edge
    _fbTrigReset   : R_TRIG;                // 复位上升沿（Reset rising edge）/ Reset rising edge
    _fbTonPress    : TON;                   // 升压段定时（Pressurise timer）/ Pressurise timer
    _fbTonStab     : TON;                   // 稳压段定时（Stabilise timer）/ Stabilise timer
    _fbTonStabExt  : TON;                   // 稳压延长定时（Stabilise extension timer）/ Stabilise extension timer
    _fbTonMeas     : TON;                   // 测量段定时（Measure timer）/ Measure timer
END_VAR

VAR CONSTANT
    DL_ESC_REAL_MAX   : REAL := 3.4E38;      // 单精度有限值判据幅值（Finite magnitude bound）/ Finite bound for REAL inputs
    DL_ESC_EPS        : REAL := 1.0E-6;      // 浮点防零容差（Divide-guard epsilon）/ Float divide-guard epsilon
    DL_ESC_PRESS_MAX  : REAL := 500.0;       // 压力输入域上限（Pressure input bound）[kPa] / Pressure input bound [kPa]
    DL_ESC_FLOW_MAX   : REAL := 5000.0;      // 流量输入域上限（Flow input bound）[sccm] / Flow input bound [sccm]
    DL_ESC_TEMP_MAX   : REAL := 200.0;       // 温度输入域上限（Temperature input bound）[℃] / Temperature input bound [degC]
    DL_ESC_TGT_MIN    : REAL := 1.0;         // 目标压力域下限（Target lower clamp）[kPa] / Target lower clamp [kPa]
    DL_ESC_TGT_MAX    : REAL := 100.0;       // 目标压力域上限（Target upper clamp）[kPa] / Target upper clamp [kPa]
    DL_ESC_TOL_MIN    : REAL := 0.01;        // 达压容差域下限（Tolerance lower clamp）[kPa] / Tolerance lower clamp [kPa]
    DL_ESC_TOL_MAX    : REAL := 50.0;        // 达压容差域上限（Tolerance upper clamp）[kPa] / Tolerance upper clamp [kPa]
    DL_ESC_LEAK_MAX   : REAL := 1.0E4;       // 漏率域上限（Leak limit ceiling）[sccm] / Leak limit ceiling [sccm]
    DL_ESC_RISE_MIN   : REAL := 0.01;        // 升压速率基准下限（Rate reference lower clamp）[kPa/s] / Rate reference lower clamp [kPa/s]
    DL_ESC_RISE_MAX   : REAL := 100.0;       // 升压速率基准上限（Rate reference upper clamp）[kPa/s] / Rate reference upper clamp [kPa/s]
    DL_ESC_COEF_MIN   : REAL := -0.05;       // 温漂系数域下限（Coefficient lower clamp）[1/K] / Coefficient lower clamp [1/K]
    DL_ESC_COEF_MAX   : REAL := 0.05;        // 温漂系数域上限（Coefficient upper clamp）[1/K] / Coefficient upper clamp [1/K]
    DL_ESC_STAB_MIN   : REAL := 0.001;       // 稳压容差域下限（Stabilisation tolerance lower clamp）[kPa] / Tolerance lower clamp [kPa]
    DL_ESC_STAB_MAX   : REAL := 50.0;        // 稳压容差域上限（Stabilisation tolerance upper clamp）[kPa] / Tolerance upper clamp [kPa]
    DL_ESC_RISE_LOWR  : REAL := 0.02;        // 供气异常判据：基准速率的 2 %（Suppy-fault ratio）[-] / Supply-fault ratio
    DL_ESC_RISE_WAIT  : REAL := 1.0;         // 升压速率判据等待秒值（Rate-test wait）[s] / Rate-test wait [s]
    DL_ESC_DTK_MIN    : REAL := 1.0;         // 温漂修正启用温差（Correction-enable temperature change）[K] / Correction-enable delta-T [K]
    DL_ESC_MS_SCALE   : REAL := 1000.0;      // 毫秒→秒换算（Milliseconds-to-seconds scale）[-] / Milliseconds-to-seconds scale
    DL_ESC_LEAK_K     : REAL := 1500.0;      // 压降率→漏率标定系数（Decay-to-leak calibration）[sccm/(kPa/s)]，偏离留档③ / Calibration constant
    DL_ESC_SCCM_MAX   : REAL := 1.0E5;       // 漏率出口上限（Leak output ceiling）[sccm] / Leak output ceiling [sccm]
    DL_ESC_DECAY_MAX  : REAL := 1.0E3;       // 压降率出口夹域（Decay output clamp）[kPa/s] / Decay output clamp [kPa/s]
    DL_ESC_ERR_PRESS  : UDINT := 16#0005_02F6; // 0005_02F6 升压超时或供气异常【故障级】/ Pressurisation failed, fault level
    DL_ESC_ERR_RISE   : UDINT := 16#0005_02F7; // 0005_02F7 测量段压力上升（源侧串漏或阀未关）【故障级】/ Pressure rising in the measure phase
    DL_ESC_ERR_STATE  : UDINT := 16#0005_02F8; // 0005_02F8 非有限输入或非法状态兜底【故障级】/ Non-finite input or illegal state fallback
    DL_ESC_INFO_EXT   : UDINT := 16#0005_01C8; // 0005_01C8 稳压未达判据已延长一次【信息级】/ Stabilisation extended once, info level
    DL_ESC_INFO_TCORR : UDINT := 16#0005_01C9; // 0005_01C9 温漂修正已启用【信息级】/ Temperature correction active, info level
    DL_ESC_INFO_WARN  : UDINT := 16#0005_01CA; // 0005_01CA 漏率落在 Warn 带【信息级】/ Leak rate inside the warn band, info level
END_VAR

// ============================================================================
// 段 1｜实例无条件周期刷新（R7/0.5：严禁置于 IF / CASE 分支内）
//      Unconditional per-cycle refresh of every instance (R7/0.5)
// ============================================================================
_fbTrigStart(CLK := bStart);                    // 启动上升沿（Start rising edge）
_bStartReq := _fbTrigStart.Q AND (NOT _bStartConsumed);   // 单拍启动请求（R25 置位点）
_fbTrigReset(CLK := bReset);                    // 复位上升沿（Reset rising edge）
_bResetEdge := _fbTrigReset.Q;                  // 复位单拍标志紧随实例赋值（R25 自清点）

// 三段各一个 TON，IN 串「段断输入标志」（R40 合规指纹：绝不跨段恒真）
// One timer per segment with the segment break folded into IN (R40)
_fbTonPress(
    IN := (_ePhase = E_DL_EscLeakPhase.ePressurize) AND (NOT _bPressBreak),
    PT := tPressurizeMax
);                                              // 升压段超时（Pressurise timeout）
_fbTonStab(
    IN := (_ePhase = E_DL_EscLeakPhase.eStabilize) AND (NOT _bStabBreak),
    PT := tStabilize
);                                              // 稳压段时长（Stabilise duration）
_fbTonStabExt(
    IN := (_ePhase = E_DL_EscLeakPhase.eStabilize) AND _bStabExtended AND (NOT _bStabExtBreak),
    PT := tStabilize
);                                              // 稳压延长段时长（Stabilise extension duration）
_fbTonMeas(
    IN := (_ePhase = E_DL_EscLeakPhase.eMeasure) AND (NOT _bMeasBreak),
    PT := tMeasure
);                                              // 测量段时长（Measure duration）

// 本拍码与条件预置（每拍重算；故障码以上拍锁存续用）
// Per-scan preset of codes and conditions, the fault code is carried from the latch
_uFaultCode := _uFaultLatched;                  // 故障码续用（Carry the latched fault code）
_uInfoCode  := 16#0000_0000;                    // 信息级码预清零（Info code preset to zero）
_bFaultCond := FALSE;                           // 故障条件预清零（Fault condition preset FALSE）

// 启动消费标志解除：输入回落即允许下一周期（R25 生命周期闭环）
// Release the start consumption flag once the input falls
IF NOT bStart THEN
    _bStartConsumed := FALSE;                   // 允许下一次上升沿（Next rising edge accepted）
END_IF

// ============================================================================
// 段 2｜断输入拍自清 + 复位通道（R40 自清 / R39 前置）
//      Segment break self-clear and the reset path, both before CASE
// ============================================================================
IF _bPressBreak THEN
    _bPressBreak := FALSE;                      // 升压段断输入拍自清（Pressurise break self-cleared）
END_IF
IF _bStabBreak THEN
    _bStabBreak := FALSE;                       // 稳压段断输入拍自清（Stabilise break self-cleared）
END_IF
IF _bStabExtBreak THEN
    _bStabExtBreak := FALSE;                    // 稳压延长断输入拍自清（Extension break self-cleared）
END_IF
IF _bMeasBreak THEN
    _bMeasBreak := FALSE;                       // 测量段断输入拍自清（Measure break self-cleared）
END_IF

IF _bResetEdge THEN
    _bDoneLatched  := FALSE;                    // 完成锁存清除（Done latch cleared）
    _bPassLatched  := FALSE;                    // 合格锁存清除（Pass latch cleared）
    _eResultHeld   := E_DL_LeakResult.eAborted; // 结果回「无结论」（Result back to the no-conclusion value）
    _fLeakHeld     := 0.0;                      // 漏率保持值清零（Held leak rate cleared）
    _fDecayHeld    := 0.0;                      // 压降率保持值清零（Held decay rate cleared）
    _bStabExtended := FALSE;                    // 延长标志清除（Extension flag cleared）
    _bStabWeak     := FALSE;                    // 弱稳定标志清除（Weak settle flag cleared）
    _nTestInt      := UDINT#0;                  // 检测计数清零（Test counter cleared）
    _nNgInt        := UDINT#0;                  // 不合格计数清零（Reject counter cleared）
    _uFaultLatched := 16#0000_0000;             // 故障码锁存清除（Latched fault code cleared）
    _uFaultCode    := 16#0000_0000;             // 本拍故障码清空，防止段7 重新锁存旧码（Clear this scan code）
    IF _ePhase = E_DL_EscLeakPhase.eFault THEN
        _ePhase := E_DL_EscLeakPhase.eIdle;     // 故障态回空闲（Fault phase back to idle）
        _bFaultCond := FALSE;                   // 故障条件清除（Fault condition cleared）
    END_IF
END_IF

// ============================================================================
// 段 3｜输入防御与参数钳位（先判可用再算值；镜像量每拍只锁一次，R38）
//      Input defense and parameter clamping, each mirror value latched once (R38)
// ============================================================================
IF (NOT (fHePressure >= (-DL_ESC_REAL_MAX) AND fHePressure <= DL_ESC_PRESS_MAX))
OR (NOT (fHeFlow >= (-DL_ESC_REAL_MAX) AND fHeFlow <= DL_ESC_FLOW_MAX))
OR (NOT (fChuckTemp >= (-DL_ESC_REAL_MAX) AND fChuckTemp <= DL_ESC_TEMP_MAX)) THEN
    _bFaultCond := TRUE;                        // 非有限或越域即故障（Non-finite or out-of-domain is a fault）
    _uFaultCode := DL_ESC_ERR_STATE;            // 0005_02F8 非有限输入【故障级】/ Non-finite input, fault level
    _fPnow   := 0.0;                            // 压力快照置零，绝不用脏值（Pressure snapshot zeroed）
    _fTnow   := 0.0;                            // 温度快照置零（Temperature snapshot zeroed）
    _fFlowNow := 0.0;                           // 流量快照置零（Flow snapshot zeroed）
ELSE
    _fPnow   := fHePressure;                    // 压力快照锁定（Pressure snapshot latched）
    _fTnow   := fChuckTemp;                     // 温度快照锁定（Temperature snapshot latched）
    _fFlowNow := fHeFlow;                       // 流量快照锁定（Flow snapshot latched）
END_IF

// 参数域钳位（R35：守卫、封顶与判据同向）
// Parameter clamping so that guard, ceiling and comparison stay in step (R35)
_fTargetEff  := LIMIT(DL_ESC_TGT_MIN, fPressTarget, DL_ESC_TGT_MAX);     // 目标压力 1~100 kPa（Target clamped）
_fTolEff     := LIMIT(DL_ESC_TOL_MIN, fPressTol, DL_ESC_TOL_MAX);        // 达压容差 0.01~50 kPa（Tolerance clamped）
_fWarnEff    := LIMIT(0.0, fLeakWarn, DL_ESC_LEAK_MAX);                  // Warn 阈 0~1E4（Warn limit clamped）
_fNgEff      := LIMIT(0.0, fLeakNg, DL_ESC_LEAK_MAX);                    // NG 阈 0~1E4（Reject limit clamped）
IF _fNgEff < _fWarnEff THEN
    _fNgEff := _fWarnEff;                       // NG 阈不得低于 Warn 阈（Reject limit never below the warn limit）
END_IF
_fRiseRefEff := LIMIT(DL_ESC_RISE_MIN, fPressRiseMax, DL_ESC_RISE_MAX);  // 升压速率基准 0.01~100（Rate reference clamped）
_fCoeffEff   := LIMIT(DL_ESC_COEF_MIN, fTempCoeff, DL_ESC_COEF_MAX);     // 温漂系数 ±0.05（Coefficient clamped）
_fStabTolEff := LIMIT(DL_ESC_STAB_MIN, fStabTol, DL_ESC_STAB_MAX);       // 稳压容差 0.001~50（Stabilise tolerance clamped）

// ============================================================================
// 段 4｜启动沿受理（R24/R25：单拍消费，消费拍与转出拍分离）
//      Start edge acceptance, single-scan consumption (R24/R25)
// ============================================================================
IF _bStartReq AND (NOT _bStartConsumed) AND bEnable AND (NOT _bFaultCond)
AND ((_ePhase = E_DL_EscLeakPhase.eIdle) OR (_ePhase = E_DL_EscLeakPhase.eVerdict)) THEN
    _bStartConsumed := TRUE;                    // 消费启动沿（Start edge consumed）
    _bDoneLatched   := FALSE;                   // 上一次完成标志清除（Previous done cleared）
    _bPassLatched   := FALSE;                   // 上一次合格标志清除（Previous pass cleared）
    _bStabExtended  := FALSE;                   // 延长标志清零（Extension flag cleared）
    _bStabWeak      := FALSE;                   // 弱稳定标志清零（Weak settle cleared）
    _fP0            := _fPnow;                  // 升压起点压力（Pressurise start pressure）
    _fStabMin       := _fPnow;                  // 稳压极值初值（Stabilise extremes seeded）
    _fStabMax       := _fPnow;                  // 稳压极大初值（Stabilise maximum seeded）
    _uInfoCode      := 16#0000_0000;            // 新一次检测起点清信息码（R44：清码点绑定新周期）
    _ePhase         := E_DL_EscLeakPhase.ePressurize;   // 进升压段（Enter pressurise）
    _bPressBreak    := TRUE;                    // 断输入一拍，三段计时都从 0 起（R40/R41）
END_IF

// ============================================================================
// 段 5｜相位状态机（ENUM + CASE，含 ELSE 非法状态兜底）
//      Phase state machine with an explicit ELSE fallback
// ============================================================================
IF _bFaultCond THEN
    _ePhase := E_DL_EscLeakPhase.eFault;        // 故障条件优先于状态机（Fault outranks the machine）
END_IF

// 掉使能冻结分支：显式排除故障态（R39 合法写法①），复位通道仍可从故障态退出
// Disable branch explicitly excludes the fault state so the reset path still works
IF (NOT bEnable) AND (_ePhase <> E_DL_EscLeakPhase.eFault) THEN
    IF (_ePhase = E_DL_EscLeakPhase.ePressurize) OR (_ePhase = E_DL_EscLeakPhase.eStabilize)
    OR (_ePhase = E_DL_EscLeakPhase.eMeasure) THEN
        _eResultHeld := E_DL_LeakResult.eAborted;   // 中止：无结论（Aborted, no conclusion）
        _bDoneLatched := TRUE;                  // 完成标志保持（Done held, per V4）
        _bPassLatched := FALSE;                 // 合格标志强制假（Pass forced FALSE）
    END_IF
    _ePhase := E_DL_EscLeakPhase.eIdle;         // 回空闲（Back to idle）
END_IF

CASE _ePhase OF

    E_DL_EscLeakPhase.eIdle: // 空闲：启动受理已在段4 完成
        // 启动动作在 CASE 之前完成（R39 前置纪律），此处保留空标签与原因注释（R31）
        // Start acceptance happens before CASE, so this label stays empty (R31)

    E_DL_EscLeakPhase.ePressurize: // 升压：等达压 / 供气异常 / 超时
        _fEtSec := TIME_TO_REAL(_fbTonPress.ET) / DL_ESC_MS_SCALE;   // 已历秒值（Elapsed seconds）
        IF ABS(_fPnow - _fTargetEff) <= _fTolEff THEN
            _ePhase      := E_DL_EscLeakPhase.eStabilize;   // 达压进稳压（Target reached, stabilise）
            _fStabMin    := _fPnow;             // 稳压极值重装（Extremes reloaded）
            _fStabMax    := _fPnow;             // 稳压极大重装（Maximum reloaded）
            _bStabBreak  := TRUE;               // 稳压定时断输入一拍（R40）
        ELSIF _fEtSec > DL_ESC_EPS THEN
            _fRiseRate := (_fPnow - _fP0) / _fEtSec;            // 升压速率（Pressurise rate）
            IF (_fRiseRate < (_fRiseRefEff * DL_ESC_RISE_LOWR))
            AND (_fEtSec > DL_ESC_RISE_WAIT) THEN
                _bFaultCond := TRUE;            // 供气异常：速率长期低于基准 2 %（Supply fault）
                _uFaultCode := DL_ESC_ERR_PRESS;    // 0005_02F6 供气异常【故障级】/ Supply fault, fault level
                _ePhase     := E_DL_EscLeakPhase.eFault;
            END_IF
        END_IF
        IF _fbTonPress.Q AND (_ePhase = E_DL_EscLeakPhase.ePressurize) THEN
            _bFaultCond := TRUE;                // 升压超时（Pressurise timeout）
            _uFaultCode := DL_ESC_ERR_PRESS;    // 0005_02F6 升压超时【故障级】/ Pressurise timeout, fault level
            _ePhase     := E_DL_EscLeakPhase.eFault;
        END_IF

    E_DL_EscLeakPhase.eStabilize: // 稳压：跟踪极差，到时判稳定
        IF _fPnow < _fStabMin THEN
            _fStabMin := _fPnow;                // 稳压极小（Stabilise minimum）
        END_IF
        IF _fPnow > _fStabMax THEN
            _fStabMax := _fPnow;                // 稳压极大（Stabilise maximum）
        END_IF
        _fStabRange := _fStabMax - _fStabMin;   // 稳压极差（Stabilise range）
        IF _bStabExtended THEN
            // 延长窗：只由延长定时器到点裁决；主稳压定时器的 Q 在延长窗内保持 TRUE，
            // 绝不能再参与裁决（否则延长置位次拍即被提前判不稳，v1.0.1 修复 D-C4-1）
            //     Extension window: arbitrated only by the extension timer (v1.0.1 fix)
            IF _fbTonStabExt.Q THEN
                IF _fStabRange <= _fStabTolEff THEN
                    _ePhase   := E_DL_EscLeakPhase.eMeasure;    // 延长后收敛：正常进测量（Settled after extension）
                    _bStabWeak := FALSE;            // 已收敛不留弱稳定标记（Settled, weak flag cleared）
                    _fPm      := _fPnow;            // 测量起点压力（Measure start pressure）
                    _fTm      := _fTnow;            // 测量起点温度（Measure start temperature）
                    _bMeasBreak := TRUE;            // 测量定时断输入一拍（R40）
                ELSE
                    _ePhase    := E_DL_EscLeakPhase.eMeasure;   // 延长后仍不稳：进测量但降级判（Deviation 4）
                    _bStabWeak := TRUE;             // 弱稳定标记（Weak settle flagged）
                    _fPm       := _fPnow;           // 测量起点压力（Measure start pressure）
                    _fTm       := _fTnow;           // 测量起点温度（Measure start temperature）
                    _bMeasBreak := TRUE;            // 测量定时断输入一拍（R40）
                END_IF
            END_IF
        ELSIF _fbTonStab.Q THEN
            IF _fStabRange <= _fStabTolEff THEN
                _ePhase   := E_DL_EscLeakPhase.eMeasure;    // 稳定判据通过进测量（Settled, measure）
                _fPm      := _fPnow;            // 测量起点压力（Measure start pressure）
                _fTm      := _fTnow;            // 测量起点温度（Measure start temperature）
                _bMeasBreak := TRUE;            // 测量定时断输入一拍（R40）
            ELSE
                _bStabExtended  := TRUE;        // 仅延长一次（Extend exactly once）
                _bStabExtBreak  := TRUE;        // 延长段定时断输入一拍（R40）
                _uInfoCode      := DL_ESC_INFO_EXT; // 0005_01C8 稳压未达判据已延长一次【信息级】/ Stabilisation extended
            END_IF
        END_IF

    E_DL_EscLeakPhase.eMeasure: // 测量：隔离窗到期结算压降与漏率
        IF _fbTonMeas.Q THEN
            _fMeasSec := TIME_TO_REAL(_fbTonMeas.ET) / DL_ESC_MS_SCALE;     // 实际测量秒值（Measured seconds）
            _fDecay   := _fPm - _fPnow;         // 压降量，有符号（Pressure drop, signed）
            IF _fDecay < 0.0 THEN
                _bFaultCond := TRUE;            // 压力上升：方向反（Pressure rising, direction reversed）
                _uFaultCode := DL_ESC_ERR_RISE; // 0005_02F7 氦源串漏或阀未关【故障级】/ Rising pressure, fault level
                _ePhase     := E_DL_EscLeakPhase.eFault;
            ELSIF _fMeasSec > DL_ESC_EPS THEN
                // 温漂修正：ΔP_corr = ΔP − P·α·ΔT（一阶线性近似，对外声明适用域）
                //     Drift correction: first-order linear approximation
                _fDtKelvin := _fTnow - _fTm;    // 测量段温差（Temperature change）
                IF (ABS(_fCoeffEff) > DL_ESC_EPS) AND (ABS(_fDtKelvin) > DL_ESC_DTK_MIN) THEN
                    _fDecayCorr := _fDecay - (_fPm * _fCoeffEff * _fDtKelvin);  // 修正后压降（Corrected drop）
                    _uInfoCode  := DL_ESC_INFO_TCORR;   // 0005_01C9 温漂修正已启用【信息级】/ Correction active
                ELSE
                    _fDecayCorr := _fDecay;     // 未启用修正（Correction not applied）
                END_IF
                IF _fDecayCorr < 0.0 THEN
                    _fDecayCorr := 0.0;         // 修正后回负按 0（Corrected drop floored to zero）
                END_IF
                _fDecayRate  := _fDecayCorr / _fMeasSec;                // 压降率（Decay rate）
                _fLeakCalc   := _fDecayRate * DL_ESC_LEAK_K;            // 漏率换算（Leak rate conversion）
                _fLeakHeld   := LIMIT(0.0, _fLeakCalc, DL_ESC_SCCM_MAX);    // 漏率夹进非负（Leak clamped）
                _fDecayHeld  := LIMIT(-DL_ESC_DECAY_MAX, _fDecayRate, DL_ESC_DECAY_MAX); // 压降率夹域（Decay clamped）

                // 三级判定：Warn 带 / NG / OK，并做流量交叉校验
                //     Three-level verdict plus the flow cross check
                IF _fLeakHeld > _fNgEff THEN
                    _eResultCalc := E_DL_LeakResult.eNg;            // 超 NG 阈（Above the reject limit）
                ELSIF _fLeakHeld > _fWarnEff THEN
                    _eResultCalc := E_DL_LeakResult.eWarn;          // 落在 Warn 带（Inside the warn band）
                    _uInfoCode   := DL_ESC_INFO_WARN;               // 0005_01CA 漏率落在 Warn 带【信息级】/ Inside the warn band
                ELSE
                    _eResultCalc := E_DL_LeakResult.eOk;            // 合格（OK）
                END_IF
                IF (_fFlowNow > _fNgEff) AND (_fLeakHeld <= _fWarnEff) THEN
                    _eResultCalc := E_DL_LeakResult.eWarn;          // 流量与换算值矛盾：至少 Warn（Corroboration mismatch）
                    _uInfoCode   := DL_ESC_INFO_WARN;               // 0005_01CA 交叉校验不一致【信息级】/ Cross check mismatch
                END_IF
                IF _bStabWeak AND (_eResultCalc = E_DL_LeakResult.eOk) THEN
                    _eResultCalc := E_DL_LeakResult.eWarn;          // 稳定判据欠佳：OK 降为 Warn（Weak settle degrades OK）
                    _uInfoCode   := DL_ESC_INFO_WARN;               // 0005_01CA 稳定判据欠佳【信息级】/ Weak settle, info level
                END_IF

                _eResultHeld  := _eResultCalc;                      // 结果锁存（Result latched）
                _bPassLatched := (_eResultCalc = E_DL_LeakResult.eOk);  // 合格锁存（Pass latched）
                _bDoneLatched := TRUE;                              // 完成锁存（Done latched）
                _nTestInt     := _nTestInt + UDINT#1;               // 检测计数 +1（Test counted）
                IF _eResultCalc = E_DL_LeakResult.eNg THEN
                    _nNgInt := _nNgInt + UDINT#1;                   // 不合格计数 +1（Reject counted）
                END_IF
                _ePhase := E_DL_EscLeakPhase.eVerdict;              // 进判定相（Enter the verdict phase）
            END_IF
        END_IF

    E_DL_EscLeakPhase.eVerdict: // 判定：结论已在测量段结算，本相只做回空闲
        _ePhase := E_DL_EscLeakPhase.eIdle;     // 结算完成回空闲（Settled, back to idle）
        _bDoneLatched := TRUE;                  // 完成标志逐拍保持（Done held, R27）

    E_DL_EscLeakPhase.eFault: // 故障：等复位沿（段2）
        // 复位通道位于 CASE 之前，此分支无需动作（R39）
        // The reset path sits before CASE, so no action is needed here (R39)

    ELSE // 兜底：非法状态
        _uFaultCode := DL_ESC_ERR_STATE;        // 0005_02F8 非法状态兜底【故障级】/ Illegal state fallback
        _bFaultCond := TRUE;                    // 置故障条件（Raise the fault condition）
        _ePhase     := E_DL_EscLeakPhase.eFault;    // 强制回故障态（Force the fault state）
END_CASE

// ============================================================================
// 段 7｜码位单一优先级链（全拍只写一次，信息级不置 bError）
//      Single priority chain for the codes, written once per scan
// ============================================================================
IF _uFaultCode <> 16#0000_0000 THEN
    _uFaultLatched := _uFaultCode;              // 故障码锁存（Latched until reset）
    uErrorId  := _uFaultCode;                   // 故障级码优先（Fault-level code wins）
    uDiagCode := _uFaultCode;                   // 诊断码同源（Diagnostic code mirrors the fault）
    bError    := TRUE;                          // 故障标志置位（Error flag raised）
ELSIF _uInfoCode <> 16#0000_0000 THEN
    uErrorId  := 16#0000_0000;                  // 信息级不占故障码（Info level leaves the fault code empty）
    uDiagCode := _uInfoCode;                    // 诊断码取信息级码（Diagnostic code takes the info code）
    bError    := FALSE;                         // 信息级不置故障位（Info level never raises the error flag）
ELSE
    uErrorId  := 16#0000_0000;                  // 无码（No code）
    uDiagCode := 16#0000_0000;                  // 无码（No code）
    bError    := FALSE;                         // 无故障（No error）
END_IF

// ============================================================================
// 段 8｜出口钳位与保持语义重写（R27/R43：结论逐拍重写，每条路径一次钳位）
//      Output clamping and held-semantics rewrite (R27/R43)
// ============================================================================
fLeakRate   := LIMIT(0.0, _fLeakHeld, DL_ESC_SCCM_MAX);                          // 漏率非负夹域（Leak clamped non-negative）
fPressDecay := LIMIT(-DL_ESC_DECAY_MAX, _fDecayHeld, DL_ESC_DECAY_MAX);          // 压降率夹域（Decay clamped）
eResult     := _eResultHeld;                                                    // 结果逐拍重写（Result rewritten every scan）
bDone       := _bDoneLatched;                                                   // 完成位逐拍重写（Done rewritten every scan）
bPass       := _bPassLatched;                                                   // 合格位逐拍重写（Pass rewritten every scan）
nTestCount  := _nTestInt;                                                       // 检测计数逐拍重写（Test counter rewritten）
nNgCount    := _nNgInt;                                                         // 不合格计数逐拍重写（Reject counter rewritten）

// 健康态仲裁（引用属主 A1 的四态语言；工件漏率 NG 不是设备健康问题）
// Health arbitration: a part leak NG is not an equipment health problem
IF _ePhase = E_DL_EscLeakPhase.eFault THEN
    eHealth := E_DL_Ne107Status.eFailure;       // 故障：供气/阀件/传感器不可信（Failure）
ELSIF NOT bEnable THEN
    eHealth := E_DL_Ne107Status.eUnknown;       // 未知：未使能（Unknown）
ELSIF (_eResultHeld = E_DL_LeakResult.eWarn) OR _bStabWeak THEN
    eHealth := E_DL_Ne107Status.eMaintenanceReq;    // 需维护：漏率入 Warn 带或稳压欠佳（Maintenance required）
ELSIF _eResultHeld = E_DL_LeakResult.eNg THEN
    eHealth := E_DL_Ne107Status.eOk;            // 正常：NG 属工件/密封面不良，设备本身健康（OK, part-level defect）
ELSE
    eHealth := E_DL_Ne107Status.eOk;            // 正常（OK）
END_IF

END_FUNCTION_BLOCK

(* ---- FB_DL_FillPreactSelfLearn.st ---- *)
(*==============================================================================
 * 组件名称 (Component)  : FB_DL_FillPreactSelfLearn
 * 所属子库 (Sublibrary) : DL_Process ｜ 版本 (Version) : 1.0.0 ｜ 2026-11-24
 * 码位     (Code Segment): 16#0005_2180（DL_Process 段内 21xx 子带）
 * 复杂度   (Complexity) : C4
 * 兼容性   (Platform)   : CODESYS 3.5+ / TwinCAT 3 / 汇川 InoProShop / 施耐德 Machine Expert
 *                         仅依赖 IEC 61131-3 标准库（TON / R_TRIG / LIMIT / ABS / REAL_TO_LREAL /
 *                         LREAL_TO_REAL），零厂商私有库
 * 开源溯源 (Provenance) : menes97/ayran-mini-fabrika / FB_Dolum PREACT / MIT /
 *                         借鉴点：粗流 / 细流两段切换与预动作量 PREACT 自学习（下落量补偿）语义
 *                         （未复制任何实现行，按 IEC 61131-3 重写为六相状态机 + 限幅学习器）
 * 功能描述 (Function)   : 灌装预动作量自学习。一轮灌装的四相节拍：eCoarse（粗流，实际重量到达
 *                         「目标 − 预动作量」即切细流）→ eFine（细流，实际重量到达「目标 − 粗流
 *                         裕度」即停阀）→ eSettle（等称重稳定或整定窗超时）→ eLearn（按最终偏差
 *                         修正预动作量并限幅）→ eDone（单拍完成回执）→ eIdle。
 *                         **学习律**：err = 实称 − 目标；PREACT := PREACT + gain × err；结果夹在
 *                         [rPreactMin, rPreactMax]，触界置 bLearnClamped。符号自证：实称超目标
 *                         （err > 0）时粗流必须更早切细流，即 PREACT 增大，公式方向正确。
 *                         **不稳定样本纪律**：整定窗超时（信息级 41）时本轮**跳过学习**——用未收敛
 *                         的读数去修正学习值，等于把气泡 / 挂料引起的瞬时偏差写成永久偏置。
 *                         **学习资产保护**：_fPreactKg / _fMargin / _iLearnCnt 属学习资产，
 *                         bReset 与 bEnable = FALSE 均**不清**（R191 声明：只降级输出 + 清状态与
 *                         锁存）；掉电保持需上层把 rPreactKg 回写 RETENTIVE 变量，本件不持有。
 *                         **COARSE_MARGIN 口径（v1.0.0 显式留置）**：裕度自学习需要「粗流段截尾
 *                         重量」这一独立观测量，本版派单未提供该引脚；在缺少中间观测的前提下
 *                         修改裕度等于用最终偏差伪造中间偏差，故本版 rCoarseMargin 只做配置量
 *                         的域钳定输出（不走学习）。v1.1 待新增 rCoarseEndKg 引脚后立项。
 * 接口     (Interface)  : 输入 bEnable / bReset（上升沿）/ bStart / rTargetKg / rActualKg /
 *                         rCoarseMarginInit / rLearnGain / rPreactMin / rPreactMax /
 *                         tSettleTimeout / bWeightStable；
 *                         输出 eState（E_DL_FillPreactSelfLearn_State）/ bBusy / bDone / bError /
 *                         iErrCode / rPreactKg / rCoarseMargin / rLastErrKg / iLearnCnt /
 *                         bLearnClamped。
 * 状态迁移表 (State Transition Table)：
 *   ① eIdle → eCoarse：bEnable 且 bStart 且组态闸通过且无锁存；拍 N 进入 / 本拍行为：清限幅
 *      标志与稳定标志、拒收本轮样本 / 拍 N+1 转出至 eCoarse。
 *   ② eCoarse → eFine：实称 ≥ 目标 − 预动作量 − 容差（本拍事件优先，R275）；拍 N 进入 /
 *      本拍行为：相级看门狗已在 CASE 外清零 / 拍 N+1 转出至 eFine。
 *   ③ eCoarse → eIdle：bEnable = FALSE（进相前置条件消失，第二出口，R98）。
 *   ④ eFine → eSettle：实称 ≥ 目标 − 粗流裕度 − 容差；拍 N 进入 / 本拍行为：拒收本轮样本 /
 *      拍 N+1 转出至 eSettle。
 *   ⑤ eFine → eIdle：bEnable = FALSE（第二出口）。
 *   ⑥ eSettle → eLearn：bWeightStable（稳定样本）；拍 N 进入 / 本拍行为：置稳定标志 /
 *      拍 N+1 转出至 eLearn。
 *   ⑦ eSettle → eLearn：tonSettle.Q（整定窗超时，信息级 41，清稳定标志，本轮跳过学习）。
 *   ⑧ eSettle → eIdle：bEnable = FALSE（第三出口）。
 *   ⑨ eLearn → eDone：单拍学习；拍 N 进入 / 本拍行为：偏差与学习值计算、限幅、非有限拒收、
 *      计数 +1，拒绝任何相推进 / 拍 N+1 转出至 eDone。
 *   ⑩ eDone → eIdle：单拍完成回执；拍 N 进入 / 本拍行为：bDone 置单拍、拒绝重复学习 /
 *      拍 N+1 转出至 eIdle。
 *   ⑪ 任意相 → eFault：相级看门狗超时 tonPhase.Q（43）；目标重量非法（42）；称重值非有限
 *      （44）；组态参数非有限（45）；非法枚举（99）。锁存后由段 7 段尾迁移闸迁相。
 *   ⑫ eFault → eIdle：bReset 上升沿；拍 N 进入 / 本拍行为：清锁存与错误码与稳定标志，
 *      **保留** rPreactKg / rCoarseMargin / iLearnCnt / bLearnClamped / rLastErrKg / 拍 N+1
 *      转出至 eIdle。出口穷举、不滞留故障态。
 * 边界     (Boundary)   : ① 两个 TON 与一个 R_TRIG 全部在 CASE 外无条件调用（R7）；IN 均含
 *                            NOT .Q 自复位项（R188）。
 *                         ② 同拍双窗配比约束（R100）：tonPhase（PT := _tSettle）覆盖 eCoarse 与
 *                            eFine 两相、tonSettle（PT := _tSettle）覆盖 eSettle 相，两使能域互斥
 *                            不相交，故共用同一超时值无竞态；语义为「单相驻留上限」，配置时须
 *                            大于最长单相时长（粗流段通常最长）。
 *                         ③ 组态域闸全覆盖（FB51-2）：六个浮点入参 rTargetKg / rActualKg /
 *                            rCoarseMarginInit / rLearnGain / rPreactMin / rPreactMax 全部逐项
 *                            枚举，无遗漏；非有限判定用自反 x <> x 与差值自减 (x−x) <> (x−x)
 *                            双判，禁用近似阈值与 ABS(x−x) 形态（R4 / R79）。
 *                         ④ 浮点比较一律带容差（1.0E-6），无 = / <> 直接判等（自反判据除外）。
 *                         ⑤ 除零防护：本件**不产生任何除法**（学习律为乘加式）；派单要求的
 *                            「目标必须为正」以量纲闸实现（rTargetKg ≤ 0 → 故障级 42），
 *                            防止后级用 rPreactKg / rTargetKg 做比例换算时除零。
 *                         ⑥ 学习值写入前必过非有限闸（R133）：非有限结果拒收并置 44，绝不写入
 *                            保持槽，避免把 NaN 变成学习起点。
 *                         ⑦ 学习增益两级限幅（FB32-3）：越出 0.05..0.8 夹紧（不故障），
 *                            防止上位误填 5.0 造成一次学习就跳满量程。
 *                         ⑧ 零全局耦合（无 GVL / VAR_EXTERNAL / %I / %Q，R1 / R2）。
 * 码表     (Codes)      : 本件按派单指定使用小整数码。信息级（永不置 bError，可每拍重算）：
 *                         41 = 整定窗超时（按不稳定样本跳过学习）；反证：该场景下 iLearnCnt 不增、
 *                              bLearnClamped 不变，输出组合与「本轮尚未学习」完全同形，只能靠码区分。
 *                         故障级（置 bError，锁存至 bReset 沿）：
 *                         42 = 目标重量非法（≤ 0 或非有限）；反证：该场景四相阈值全部退化，
 *                              输出与「刚开始灌装」同形，必须独立成码且作为首因优先判定。
 *                         43 = 相级看门狗超时（粗流 / 细流相驻留超限）；反证：该场景实称长期不达
 *                              阈值、iLearnCnt 不增，与「慢速灌装仍在进行」输出全同形。
 *                         44 = 称重值非有限（仪表失效）；反证：与 43 的区别是「有无读数」而非
 *                              「读数是否推进」，两者补救动作不同（换仪表 / 查阀门节拍）。
 *                         45 = 组态参数非有限（裕度初值 / 学习增益 / 预动作量限幅）；反证：该类
 *                              参数是静态配置，与过程量失效的补救动作（改配方 vs 修设备）不同。
 *                         99 = 非法状态枚举值（ELSE 兜底）。
 * 分工声明 (Scope)      : 粗流阀 / 细流阀的实际开闭命令归灌装时序件（本件只输出相位，相位即
 *                         命令语义）；称重滤波与稳定判据归上游称重件（本件只接收 bWeightStable）；
 *                         配方级目标重量下发归配方管理件。本件只做**预动作量单参数学习的闭环**。
 * 归属     (Ownership)  : E_DL_FillPreactSelfLearn_State 归属本文件（全库唯一定义，R264）。
 * 命名偏离 (Naming Ex.) : 本件按派单原文保留 r 前缀表示 REAL（rTargetKg / rActualKg /
 *                         rCoarseMarginInit / rLearnGain / rPreactMin / rPreactMax / rPreactKg /
 *                         rCoarseMargin / rLastErrKg），i 前缀表示 INT（iErrCode），i 前缀表示
 *                         DINT（iLearnCnt，计数语义按 FB51-7② 归 DINT）；内部计算一律升位到
 *                         LREAL 的 f 前缀。与规范 1.2 节存在登记偏离，接口契约优先不改名。
 * 红线自检 (Redline)    : R1 ✓ 零 GVL / VAR_EXTERNAL ｜ R2 ✓ 零 %I/%Q ｜ R3 ✓ 纯 IEC 61131-3
 *                         ｜ R4 ✓ 无除法 + 浮点容差比较 + 自反/差值双判非有限 + 除零量纲闸
 *                         ｜ R5 ✓ 逐行同行中英双语注释 ｜ R6 ✓ 七态 ENUM + CASE + ELSE 兜底
 *                         ｜ R7 ✓ TON / R_TRIG 全在 CASE 外无条件调用 ｜ R8 ✓ 无 METHOD（全内联）
 *                         ｜ R10 ✓ 无构造式转换（仅 REAL_TO_LREAL / LREAL_TO_REAL）｜ R11 ✓ 声明
 *                         全分号结尾 ｜ R12 ✓ ENUM 成员用 := ｜ R14 ✓ 无 PROPERTY
 *                         ｜ R16 ✓ 不引用任何外部 FB/FC（LIMIT / ABS 为 IEC 标准函数）。
 * 修订历史 (Revision)   : 2026-11-24  v1.0.0  R81-B 首版（COARSE_MARGIN 自学习显式留置 v1.1）
 * 验收向量 (Acceptance) :
 *   V1 欠灌学习：rTargetKg=1.000、rPreactKg 初值 0.100（限幅 0.02..0.35）、rLearnGain=0.3、
 *      rCoarseMarginInit=0.050、实称 0.980 → err=-0.020、新 PREACT=0.100+0.3×(-0.020)=0.094、
 *      iLearnCnt+1、bLearnClamped=FALSE、rLastErrKg=-0.020、eState 走 eDone 后回 eIdle。
 *   V2 触界限幅：rPreactKg=0.349、实称 1.060（err=+0.060）→ 原始值 0.367 超 0.35 →
 *      rPreactKg=0.350、bLearnClamped=TRUE、iLearnCnt+1。
 *   V3 不稳定样本：bWeightStable 恒 FALSE、tSettleTimeout=T#2S → eSettle 驻留 2s 后 tonSettle.Q →
 *      eLearn、iErrCode=41、iLearnCnt 不增、rPreactKg 不变、bLearnClamped 不变、bError=FALSE。
 *   V4 目标非法：rTargetKg=0.0 → eState=eFault、iErrCode=42、bError=TRUE、bBusy=FALSE；
 *      bReset 上升沿 → eState=eIdle、bError=FALSE、rPreactKg 保持故障前值（学习资产不清）。
 *   V5 称重非有限：rActualKg 置 NaN → eState=eFault、iErrCode=44、bError=TRUE。
 *   V6 增益越域：rLearnGain=5.0 → 夹紧为 0.8（不故障，bError=FALSE），一次学习跳变量不超过
 *      0.8×err；rLearnGain=0.001 → 夹紧为 0.05。
 *   V7 粗流超时：rPreactKg 使粗流阈值极低、实称恒 0、tSettleTimeout=T#1S → eCoarse 驻留 1s 后
 *      eState=eFault、iErrCode=43、bError=TRUE。
 *============================================================================*)

(*-----------------------------------------------------------------------------
 * 枚举: E_DL_FillPreactSelfLearn_State（灌装预动作量学习相位；eFault 为安全相）
 *----------------------------------------------------------------------------*)
TYPE E_DL_FillPreactSelfLearn_State :
(
    eIdle   := 0,     // 空闲：等启动条件，学习资产保持 / Idle: waiting for the start condition, learning assets kept
    eCoarse := 10,    // 粗流相：实际重量到「目标 − 预动作量」切细流 / Coarse: switch to fine when the weight reaches the target minus PREACT
    eFine   := 20,    // 细流相：实际重量到「目标 − 粗流裕度」停阀 / Fine: close the valve at the target minus the coarse margin
    eSettle := 30,    // 整定相：等称重稳定或整定窗超时 / Settle: waiting for weight stability or the settle window
    eLearn  := 40,    // 学习相：单拍更新预动作量并限幅 / Learn: one-scan PREACT update with clamping
    eDone   := 50,    // 完成相：单拍回执 / Done: one-scan completion receipt
    eFault  := 90     // 故障安全相：锁存成因，拒绝学习推进 / Fault safe phase: latched cause, no learning progress
);
END_TYPE

FUNCTION_BLOCK FB_DL_FillPreactSelfLearn
VAR_INPUT
    bEnable       : BOOL := FALSE;          // 使能：FALSE 回空闲（学习资产保留）/ Enable, FALSE returns to idle and keeps the learning assets
    bReset        : BOOL := FALSE;          // 复位（上升沿；清锁存与状态，不清学习值）/ Reset rising edge clearing latch and phase but not the learned values
    bStart        : BOOL := FALSE;          // 启动（电平，eIdle 出口判据）/ Start level, an eIdle exit criterion
    rTargetKg     : REAL := 0.0;            // 目标灌装重量，域 > 0 且有限 [kg] / Target fill weight, positive and finite
    rActualKg     : REAL := 0.0;            // 实称重量（称重件输出）[kg] / Measured weight delivered by the weighing component
    rCoarseMarginInit : REAL := 0.05;       // 粗流裕度配置初值，钳在 0..目标/2 [kg] / Configured coarse margin, clamped to zero through half the target
    rLearnGain    : REAL := 0.3;            // 学习增益，有效域 0.05..0.8，越域夹紧 [1] / Learning gain, clamped into 0.05 through 0.8
    rPreactMin    : REAL := 0.02;           // 预动作量下限 [kg] / PREACT lower limit
    rPreactMax    : REAL := 0.35;           // 预动作量上限，须 ≥ rPreactMin [kg] / PREACT upper limit, at least the lower limit
    tSettleTimeout : TIME := T#3S;          // 单相驻留上限（整定窗 + 粗/细流看门狗），有效域 50ms..10min [s] / Per-phase dwell limit, valid domain 50 ms through 10 min
    bWeightStable : BOOL := FALSE;          // 称重稳定（称重件判据）/ Weight stable, delivered by the weighing component
END_VAR
VAR_OUTPUT
    eState        : E_DL_FillPreactSelfLearn_State;   // 当前相位出口（段 8 单点映射）/ Current phase outlet mapped once at segment 8
    bBusy         : BOOL;                   // 本轮灌装进行中 / A fill cycle in progress
    bDone         : BOOL;                   // 本轮完成单拍脉冲 / One-scan cycle completion pulse
    bError        : BOOL;                   // 故障锁存标志 / Fault latch flag
    iErrCode      : INT := 0;               // 错误码（故障期锁存回放，非故障期为信息码）/ Error code, latched in fault and the info code otherwise
    rPreactKg     : REAL := 0.0;            // 当前预动作量（学习资产，复位不清）[kg] / Current PREACT, a learning asset kept across resets
    rCoarseMargin : REAL := 0.0;            // 当前粗流裕度（本版为域钳定配置量）[kg] / Current coarse margin, a clamped configuration value in this version
    rLastErrKg    : REAL := 0.0;            // 上次偏差 = 实称 − 目标 [kg] / Last deviation, measured minus target
    iLearnCnt     : DINT := 0;              // 学习成功累计次数 [次] / Cumulative successful learning count
    bLearnClamped : BOOL;                   // 上次学习是否被限幅 / Whether the last learning was clamped
END_VAR
VAR
    _eState       : E_DL_FillPreactSelfLearn_State := E_DL_FillPreactSelfLearn_State.eIdle;   // 内部相位（CASE 唯一写入目标）/ Internal phase, the only CASE write target
    _bFaultLatch  : BOOL := FALSE;          // 故障锁存位（仅 bReset 上升沿清除）/ Fault latch bit, cleared only by the bReset rising edge
    _iErrLatch    : INT := 0;               // 锁存故障码（故障期唯一回放源，FB33-1）/ Latched fault code, the only replay source during fault
    _iInfoCode    : INT := 0;               // 信息级码（41，永不置 bError）/ Info-level code 41, never raising bError
    _iErrTmp      : INT := 0;               // 当拍故障首因中间量 / First fault cause of this scan
    _bFaultReq    : BOOL := FALSE;          // 当拍故障请求标志（段 7 统一锁存）/ Fault request of this scan latched at segment 7
    _bCfgOk       : BOOL := TRUE;           // 组态与入参闸通过标志 / Configuration and argument gate flag
    _bInit        : BOOL := FALSE;          // 首扫初始化已执行标志（学习起点，FB50-2）/ First-scan initialisation flag for the learning start point
    _bDonePulse   : BOOL := FALSE;          // 完成内部单拍位（段 1 预置，段 8 映射）/ Internal one-scan done bit preset at segment 1
    _bSettledStable : BOOL := FALSE;        // 本轮样本稳定标志（稳定才学习）/ Stability flag of this cycle, learning happens only when stable
    _bLearnClamped : BOOL := FALSE;         // 上次学习限幅标志（内部保持量）/ Clamp flag of the last learning, an internal holding value
    _fTarget      : LREAL := 0.0;           // 目标重量升位副本 [kg] / Promoted copy of the target weight
    _fActual      : LREAL := 0.0;           // 实称重量升位副本 [kg] / Promoted copy of the measured weight
    _fMarginInit  : LREAL := 0.0;           // 粗流裕度初值升位副本 [kg] / Promoted copy of the configured coarse margin
    _fGainRaw     : LREAL := 0.0;           // 学习增益升位副本（未夹紧）[1] / Promoted learning gain before clamping
    _fGain        : LREAL := 0.0;           // 学习增益夹紧值 [1] / Clamped learning gain
    _fPmin        : LREAL := 0.0;           // 预动作量有效下限（钳后）[kg] / Effective PREACT lower limit after clamping
    _fPmax        : LREAL := 0.0;           // 预动作量有效上限（钳后）[kg] / Effective PREACT upper limit after clamping
    _fPreactKg    : LREAL := 0.0;           // 预动作量学习值（学习资产，复位不清）[kg] / Learned PREACT kept across resets
    _fMargin      : LREAL := 0.0;           // 粗流裕度派生量（每拍由初值域钳定）[kg] / Derived coarse margin clamped from the initial value each scan
    _fLastErr     : LREAL := 0.0;           // 上次偏差保持量 [kg] / Holding value of the last deviation
    _fErr         : LREAL := 0.0;           // 本轮偏差临时量 [kg] / Temporary deviation of this cycle
    _fRaw         : LREAL := 0.0;           // 学习原始结果（夹紧前）[kg] / Raw learning result before clamping
    _fClamped     : LREAL := 0.0;           // 学习夹紧后结果 [kg] / Learning result after clamping
    _iLearnCnt    : DINT := 0;              // 学习成功次数（学习资产，复位不清）[次] / Successful learning count kept across resets
    _tSettle      : TIME := T#3S;           // 单相驻留上限钳定值（两级回退结果）[s] / Clamped per-phase dwell limit after the two-level fallback
    rtReset       : R_TRIG;                 // bReset 边沿实例（段 3 无条件调用，R18）/ bReset edge instance called unconditionally
    tonPhase      : TON;                    // 粗流 / 细流相级看门狗（段 3 无条件调用）/ Phase watchdog for coarse and fine, called unconditionally
    tonSettle     : TON;                    // 整定窗计时器（段 3 无条件调用）/ Settle window timer called unconditionally
END_VAR
VAR CONSTANT
    DL_FPS_ZERO      : LREAL := 0.0;              // 浮点零基准（作有限性判据的对照量）[-] / Float zero used as the finiteness reference
    DL_FPS_EPS       : LREAL := 1.0E-6;           // 浮点比较容差（重量级 kg 下约 1 mg）[kg] / Float comparison tolerance
    DL_FPS_HALF      : LREAL := 0.5;              // 系数 0.5（中位起点与裕度上限）[1] / Factor 0.5 used for the midpoint and the margin cap
    DL_FPS_GAIN_MIN  : LREAL := 0.05;             // 学习增益下限（越界夹紧，不故障）[1] / Learning gain lower bound, clamped without fault
    DL_FPS_GAIN_MAX  : LREAL := 0.8;              // 学习增益上限（越界夹紧，不故障）[1] / Learning gain upper bound, clamped without fault
    DL_FPS_T_MIN     : TIME := T#50MS;            // 单相驻留上限下限 [s] / Per-phase dwell limit lower bound
    DL_FPS_T_MAX     : TIME := T#10M;             // 单相驻留上限上限 [s] / Per-phase dwell limit upper bound
    DL_FPS_T_DEF     : TIME := T#3S;              // 单相驻留上限默认回退值（本身在域内）[s] / Default fallback dwell limit, already inside the domain
    DL_FPS_ONE_DINT  : DINT := 1;                 // 计数步进一 [1] / Counter step of one
END_VAR

(* —— 段 1：中间量预置（只清单拍标志与扫描量，不清学习资产 / 锁存 / 稳定标志，FB32-1） —— *)
_iErrTmp    := 0;                          // 当拍故障首因复位 / Scan first fault cause reset
_bFaultReq  := FALSE;                      // 当拍故障请求复位 / Scan fault request reset
_bCfgOk     := TRUE;                       // 组态闸标志复位 / Configuration gate flag reset
_bDonePulse := FALSE;                      // 完成单拍位预置（单拍路径唯一预置点，FB51-8）/ Done pulse preset, the single preset point

(* —— 段 2：REAL 入参升位（R10 标准转换，内部一律 LREAL 运算防累积误差） —— *)
_fTarget     := REAL_TO_LREAL(rTargetKg);          // 目标重量升位 / Target weight promoted
_fActual     := REAL_TO_LREAL(rActualKg);          // 实称重量升位 / Measured weight promoted
_fMarginInit := REAL_TO_LREAL(rCoarseMarginInit);  // 裕度初值升位 / Configured margin promoted
_fGainRaw    := REAL_TO_LREAL(rLearnGain);         // 学习增益升位 / Learning gain promoted
_fPmin       := REAL_TO_LREAL(rPreactMin);         // 限幅下限升位 / PREACT lower limit promoted
_fPmax       := REAL_TO_LREAL(rPreactMax);         // 限幅上限升位 / PREACT upper limit promoted

(* —— 段 3：时间参数两级回退（越域回默认常量，默认常量在域内故无需二级钳定，FB32-3） —— *)
IF (tSettleTimeout < DL_FPS_T_MIN) OR (tSettleTimeout > DL_FPS_T_MAX) THEN
    _tSettle := DL_FPS_T_DEF;              // 越域：回一级默认常量 / Out of domain: fall back to the default constant
ELSE
    _tSettle := tSettleTimeout;            // 域内：原值采用 / Inside the domain: take the value as given
END_IF

(* —— 段 4：组态域闸全覆盖（六个浮点入参逐项枚举，FB51-2；非有限双判，R4 / R79） —— *)
IF (_fTarget <> _fTarget) OR ((_fTarget - _fTarget) <> (_fTarget - _fTarget)) THEN
    _bCfgOk  := FALSE;                     // 目标重量非有限 / Target weight is not finite
    _iErrTmp := 42;                        // 故障级：目标重量非法 / Fault: illegal target weight
END_IF
IF _bCfgOk THEN
    IF _fTarget <= DL_FPS_EPS THEN
        _bCfgOk  := FALSE;                 // 目标重量非正（量纲闸，防后级比例换算除零）/ Non-positive target, a dimensional gate against division by zero downstream
        _iErrTmp := 42;                    // 故障级：目标重量非法 / Fault: illegal target weight
    END_IF
END_IF
IF _bCfgOk THEN
    IF (_fActual <> _fActual) OR ((_fActual - _fActual) <> (_fActual - _fActual)) THEN
        _bCfgOk  := FALSE;                 // 实称重量非有限（仪表失效）/ Measured weight is not finite
        _iErrTmp := 44;                    // 故障级：称重值非有限 / Fault: non-finite measured weight
    END_IF
END_IF
IF _bCfgOk THEN
    IF ((_fMarginInit <> _fMarginInit) OR ((_fMarginInit - _fMarginInit) <> (_fMarginInit - _fMarginInit)))
        OR ((_fGainRaw <> _fGainRaw) OR ((_fGainRaw - _fGainRaw) <> (_fGainRaw - _fGainRaw)))
        OR ((_fPmin <> _fPmin) OR ((_fPmin - _fPmin) <> (_fPmin - _fPmin)))
        OR ((_fPmax <> _fPmax) OR ((_fPmax - _fPmax) <> (_fPmax - _fPmax))) THEN
        _bCfgOk  := FALSE;                 // 组态参数非有限 / A configuration parameter is not finite
        _iErrTmp := 45;                    // 故障级：组态参数非有限 / Fault: non-finite configuration parameter
    END_IF
END_IF

(* —— 段 5：参数夹紧与有效限幅（增益夹紧不故障；限幅倒置两级回退，FB32-3） —— *)
_fGain := LIMIT(DL_FPS_GAIN_MIN, _fGainRaw, DL_FPS_GAIN_MAX);   // 学习增益夹紧到 0.05..0.8 / Gain clamped into 0.05 through 0.8
IF _fPmin < DL_FPS_ZERO THEN
    _fPmin := DL_FPS_ZERO;                 // 预动作量下限不得为负（负值等于反向补偿）/ PREACT lower limit forced non-negative
END_IF
IF _fPmin > _fPmax THEN
    _fPmin := DL_FPS_ZERO;                 // 限幅倒置一级回退：下限回零 / Inverted limits fall back to a zero lower bound
    _fPmax := _fTarget * DL_FPS_HALF;      // 限幅倒置二级回退：上限按目标半量钳定（域几何内点）/ Upper bound clamped to half the target
END_IF
IF _fTarget > DL_FPS_EPS THEN
    _fMargin := LIMIT(DL_FPS_ZERO, _fMarginInit, _fTarget * DL_FPS_HALF);   // 裕度钳在 0..目标/2，防裕度过大导致细流段根本不进 / Margin clamped to avoid skipping the fine phase
ELSE
    _fMargin := DL_FPS_ZERO;               // 目标非法时裕度归零（等待段 4 的 42 锁存接管）/ Margin zeroed while the illegal target is latched
END_IF

(* —— 段 6：首扫学习起点初始化（组态闸通过后才执行，FB50-2①；复位沿**不**重跑，学习资产保留） —— *)
IF (NOT _bInit) AND _bCfgOk THEN
    _bInit     := TRUE;                                        // 置首扫完成标志 / Mark the first scan done
    _fPreactKg := (_fPmin + _fPmax) * DL_FPS_HALF;             // 起点取限幅中位（在限幅内且非零，减少首轮偏差）/ Start at the limit midpoint, inside the limits and non-zero
    _fLastErr  := DL_FPS_ZERO;                                 // 偏差保持量归零 / Deviation holding value zeroed
    _iLearnCnt := 0;                                           // 学习计数归零 / Counter zeroed
END_IF

(* —— 段 7：边沿与定时器（CASE 外无条件调用，R7；IN 均含 NOT .Q 自复位，R188） —— *)
rtReset(CLK := bReset);                    // bReset 边沿无条件刷新（R18）/ bReset edge refreshed unconditionally
tonPhase(IN := ((_eState = E_DL_FillPreactSelfLearn_State.eCoarse)
                OR (_eState = E_DL_FillPreactSelfLearn_State.eFine))
               AND (NOT tonPhase.Q) AND (NOT _bFaultLatch),
         PT := _tSettle);                  // 粗流 / 细流相级看门狗（使能域与 tonSettle 互斥）/ Phase watchdog with a domain disjoint from tonSettle
tonSettle(IN := (_eState = E_DL_FillPreactSelfLearn_State.eSettle) AND (NOT tonSettle.Q) AND (NOT _bFaultLatch),
          PT := _tSettle);                 // 整定窗计时 / Settle window timer

(* —— 段 8：状态机主体（唯一相位写入点；故障只置请求，锁存与迁相由段 9 执行，R21） —— *)
CASE _eState OF
    E_DL_FillPreactSelfLearn_State.eIdle :
        (* 迁移①：启动条件成立进粗流相 *)
        IF bEnable AND bStart AND _bCfgOk AND (NOT _bFaultLatch) THEN
            _bSettledStable := FALSE;                                 // 本轮样本稳定标志复位 / Stability flag of this cycle cleared
            _bLearnClamped  := FALSE;                                 // 本轮限幅标志复位（学习资产本身不动）/ Clamp flag of this cycle cleared, the learned value itself is kept
            _iInfoCode      := 0;                                     // 信息码复位 / Info code cleared
            _eState         := E_DL_FillPreactSelfLearn_State.eCoarse;   // 进粗流相 / Move to the coarse phase
        END_IF

    E_DL_FillPreactSelfLearn_State.eCoarse :
        (* 迁移②：实称到达「目标 − 预动作量」即切细流（本拍事件优先于超时，R275） *)
        IF _fActual >= ((_fTarget - _fPreactKg) - DL_FPS_EPS) THEN
            _eState := E_DL_FillPreactSelfLearn_State.eFine;          // 切细流 / Switch to the fine phase
        ELSIF NOT bEnable THEN
            _eState := E_DL_FillPreactSelfLearn_State.eIdle;          // 迁移③：前置条件消失回空闲 / Precondition gone, back to idle
        END_IF

    E_DL_FillPreactSelfLearn_State.eFine :
        (* 迁移④：实称到达「目标 − 粗流裕度」即停阀进整定 *)
        IF _fActual >= ((_fTarget - _fMargin) - DL_FPS_EPS) THEN
            _eState := E_DL_FillPreactSelfLearn_State.eSettle;        // 进整定相 / Move to settle
        ELSIF NOT bEnable THEN
            _eState := E_DL_FillPreactSelfLearn_State.eIdle;          // 迁移⑤：前置条件消失回空闲 / Precondition gone, back to idle
        END_IF

    E_DL_FillPreactSelfLearn_State.eSettle :
        (* 迁移⑥/⑦/⑧：稳定样本、整定超时（跳过学习）、失能三出口（R98 出口 ≥ 2） *)
        IF bWeightStable THEN
            _bSettledStable := TRUE;                                  // 稳定样本：允许学习 / Stable sample, learning allowed
            _eState := E_DL_FillPreactSelfLearn_State.eLearn;         // 迁移⑥：进学习相 / Move to learn
        ELSIF tonSettle.Q THEN
            _bSettledStable := FALSE;                                 // 不稳定样本：本轮跳过学习 / Unstable sample, this cycle skips learning
            _iInfoCode      := 41;                                    // 信息级：整定窗超时（不置 bError）/ Info: settle window timeout, bError stays false
            _eState := E_DL_FillPreactSelfLearn_State.eLearn;         // 迁移⑦：仍进学习相以更新偏差 / Still move to learn to refresh the deviation
        ELSIF NOT bEnable THEN
            _eState := E_DL_FillPreactSelfLearn_State.eIdle;          // 迁移⑧：前置条件消失回空闲 / Precondition gone, back to idle
        END_IF

    E_DL_FillPreactSelfLearn_State.eLearn :
        (* 迁移⑨：单拍学习；拍 N 进入 / 本拍行为：偏差与学习值更新、限幅、非有限拒收 / 拍 N+1 转出至 eDone *)
        _fErr        := _fActual - _fTarget;                          // 本轮偏差 = 实称 − 目标 [kg] / Deviation of this cycle
        _fLastErr    := _fErr;                                        // 偏差保持量更新（每轮都记，含不稳定样本）/ Deviation kept every cycle including unstable samples
        (* 稳定标志在本分支只读不写（禁止自赋值死语句，R261） *)
        IF _bSettledStable THEN
            _fRaw := _fPreactKg + (_fGain * _fErr);                   // 学习律：PREACT + gain × err / Learning law
            IF (_fRaw <> _fRaw) OR ((_fRaw - _fRaw) <> (_fRaw - _fRaw)) THEN
                _iErrTmp   := 44;                                     // 故障级：学习结果非有限（保持槽拒收，R133）/ Fault: non-finite result rejected
                _bFaultReq := TRUE;                                   // 请求段 9 锁存 / Request the latch at segment 9
            ELSE
                _fClamped := LIMIT(_fPmin, _fRaw, _fPmax);             // 限幅到 [下限, 上限] / Clamped into the configured limits
                IF ABS(_fClamped - _fRaw) > DL_FPS_EPS THEN
                    _bLearnClamped := TRUE;                           // 触界：本轮学习被限幅 / Clamped this cycle
                ELSE
                    _bLearnClamped := FALSE;                          // 未触界：正常学习 / No clamping this cycle
                END_IF
                _fPreactKg := _fClamped;                              // 学习值写入（唯一写入点，已过非有限闸）/ Single write point after the finiteness gate
                _iLearnCnt := _iLearnCnt + DL_FPS_ONE_DINT;            // 学习成功计数 +1 / Successful learning count incremented
            END_IF
        END_IF
        _eState := E_DL_FillPreactSelfLearn_State.eDone;              // 迁移⑨：进完成相 / Move to done

    E_DL_FillPreactSelfLearn_State.eDone :
        (* 迁移⑩：单拍完成回执；拍 N 进入 / 本拍行为：bDone 置单拍一次，拒绝重复学习 / 拍 N+1 转出至 eIdle *)
        _bDonePulse := TRUE;                                          // 完成内部单拍置位（段 10 映射）/ Internal done pulse raised and mapped at segment 10
        _eState     := E_DL_FillPreactSelfLearn_State.eIdle;          // 回空闲相 / Back to idle

    E_DL_FillPreactSelfLearn_State.eFault :
        (* 迁移⑫：复位沿出口（唯一出口，穷举可达）；学习资产一律保留）
           拍 N 进入 / 本拍行为：清锁存、错误码、稳定标志，拒绝任何学习推进 / 拍 N+1 转出至 eIdle *)
        IF rtReset.Q THEN
            _bFaultLatch    := FALSE;                                 // 清故障锁存 / Clear the fault latch
            _iErrLatch      := 0;                                     // 清锁存故障码 / Clear the latched fault code
            _iInfoCode      := 0;                                     // 清信息码 / Clear the info code
            _bSettledStable := FALSE;                                 // 清稳定标志（避免用旧样本） / Clear the stability flag to avoid reusing an old sample
            _eState         := E_DL_FillPreactSelfLearn_State.eIdle;  // 回空闲相，不滞留故障态 / Back to idle, never parked in fault
        END_IF

ELSE
    (* 迁移⑪（枚举兜底）：非法枚举值 → 故障级 99（R6） *)
    IF NOT _bFaultLatch THEN
        _iErrLatch   := 99;                    // 故障级：非法状态枚举值 / Fault: illegal state enum value
        _bFaultLatch := TRUE;                  // 置故障锁存（码位赋值 3 行内配对，R45）/ Latch the fault within three lines
    END_IF
END_CASE

(* —— 段 9：当拍故障请求锁存（定时器超时 / 组态闸）+ 段尾迁移闸 + 撤使能降级 —— *)
IF tonPhase.Q AND (NOT _bFaultLatch) THEN
    _iErrLatch   := 43;                        // 故障级：粗流 / 细流相级看门狗超时 / Fault: coarse or fine phase watchdog timeout
    _bFaultLatch := TRUE;                      // 置故障锁存 / Latch the fault
END_IF
IF (NOT _bCfgOk) AND (NOT _bFaultLatch) THEN
    _iErrLatch   := _iErrTmp;                  // 锁存组态首因 / Latch the configuration first cause
    _bFaultLatch := TRUE;                      // 置故障锁存 / Latch the fault
END_IF
IF _bFaultReq AND (NOT _bFaultLatch) THEN
    _iErrLatch   := _iErrTmp;                  // 锁存学习结果非有限首因 / Latch the non-finite result cause
    _bFaultLatch := TRUE;                      // 置故障锁存 / Latch the fault
END_IF
IF _bFaultLatch AND (_eState <> E_DL_FillPreactSelfLearn_State.eFault) THEN
    _eState := E_DL_FillPreactSelfLearn_State.eFault;   // 锁存即迁相（段尾统一执行，FB50-1④）/ Latch forces the fault phase at the tail
END_IF
IF (NOT bEnable) AND (NOT _bFaultLatch) AND (_eState <> E_DL_FillPreactSelfLearn_State.eIdle) THEN
    _eState := E_DL_FillPreactSelfLearn_State.eIdle;    // 撤使能：回空闲（学习资产保留，R191 降级声明）/ Disable: back to idle keeping the learning assets
END_IF

(* —— 段 10：统一出口（单点映射；连续量出口再做一次非有限防护，FB51-3 / R273） —— *)
eState  := _eState;                            // 相位映射 / Phase mapping
bBusy   := (_eState = E_DL_FillPreactSelfLearn_State.eCoarse)
           OR (_eState = E_DL_FillPreactSelfLearn_State.eFine)
           OR (_eState = E_DL_FillPreactSelfLearn_State.eSettle)
           OR (_eState = E_DL_FillPreactSelfLearn_State.eLearn);   // 本轮进行中 / Cycle in progress
bDone   := _bDonePulse;                        // 完成单拍映射 / Completion pulse mapping
bError  := _bFaultLatch;                       // 故障标志取锁存位 / Fault flag taken from the latch
IF _bFaultLatch THEN
    iErrCode := _iErrLatch;                    // 故障期回放锁存码（FB33-1）/ Replay the latched code during fault
ELSE
    iErrCode := _iInfoCode;                    // 非故障期输出信息码（41 永不置 bError，R101）/ Info code outside fault, never raising bError
END_IF
IF (_fPreactKg <> _fPreactKg) OR ((_fPreactKg - _fPreactKg) <> (_fPreactKg - _fPreactKg)) THEN
    _fPreactKg := DL_FPS_ZERO;                 // 保持槽污染兜底：归零（三件套中的连续量安全侧）/ Contaminated holding value forced to zero
    rPreactKg  := 0.0;                         // 出口同步归零 / Outlet follows the guard
ELSE
    rPreactKg  := LREAL_TO_REAL(_fPreactKg);   // 学习值出口（降位为 REAL）/ Learning value outlet demoted to REAL
END_IF
IF (_fMargin <> _fMargin) OR ((_fMargin - _fMargin) <> (_fMargin - _fMargin)) THEN
    rCoarseMargin := 0.0;                      // 裕度污染兜底：归零 / Contaminated margin forced to zero
ELSE
    rCoarseMargin := LREAL_TO_REAL(_fMargin);  // 裕度出口 / Margin outlet
END_IF
IF (_fLastErr <> _fLastErr) OR ((_fLastErr - _fLastErr) <> (_fLastErr - _fLastErr)) THEN
    rLastErrKg := 0.0;                         // 偏差污染兜底：归零 / Contaminated deviation forced to zero
ELSE
    rLastErrKg := LREAL_TO_REAL(_fLastErr);    // 偏差出口 / Deviation outlet
END_IF
iLearnCnt     := _iLearnCnt;                   // 学习计数出口 / Learning count outlet
bLearnClamped := _bLearnClamped;               // 限幅标志出口 / Clamp flag outlet
END_FUNCTION_BLOCK
